(* IEC 61131-3 sources: STAR-PLC-Agent/results/raw/codex_matrix_resume_20261114/codex_deepseek/PUB012/functional/attempt_0001, 1 file *)

(* ---- test_program.st ---- *)
PROGRAM PLC_PRG
VAR
 BenchStep : UDINT := 0;
 BenchCalls : UDINT := 0;
 BenchDone : BOOL := FALSE;
 BenchLastTime : TIME := T#0ms;
 BenchClockReady : BOOL := FALSE;
 BenchCurrentTime : TIME := T#0ms;
 TraceDt : ARRAY[0..69] OF UDINT;
 BenchUut0 : FB_Task;
 BenchUut1 : FB_Task;
 BenchUut2 : FB_Task;
 BenchUut3 : FB_Task;
 BenchUut4 : FB_Task;
 BenchUut5 : FB_Task;
 BenchUut6 : FB_Task;
 BenchUut7 : FB_Task;
 TraceIn_THICKNESS_FAULT : ARRAY[0..69] OF BOOL;
 TraceIn_THICKNESS_SIGNAL_VALID : ARRAY[0..69] OF BOOL;
 TraceIn_CUTTING_RUN : ARRAY[0..69] OF BOOL;
 TraceIn_FaultTimestamp : ARRAY[0..69] OF DINT;
 TraceIn_CycleTime : ARRAY[0..69] OF TIME;
 TraceOut_THICKNESS_ALARM : ARRAY[0..69] OF BOOL;
 TraceOut_Slab_Fault_Counter : ARRAY[0..69] OF UINT;
 TraceOut_Slab_Runtime_Accumulator : ARRAY[0..69] OF LTIME;
 TraceOut_Slab_Fault_History_0 : ARRAY[0..69] OF DINT;
 TraceOut_Slab_Fault_History_1 : ARRAY[0..69] OF DINT;
 TraceOut_Slab_Fault_History_2 : ARRAY[0..69] OF DINT;
 TraceOut_Slab_Fault_History_3 : ARRAY[0..69] OF DINT;
 TraceOut_Slab_Fault_History_4 : ARRAY[0..69] OF DINT;
END_VAR

IF NOT BenchDone THEN
 BenchCurrentTime := TIME();
 IF NOT BenchClockReady THEN
  BenchLastTime := BenchCurrentTime;
  BenchClockReady := TRUE;
 ELSE
 CASE BenchStep OF
 0:
  IF BenchCurrentTime - BenchLastTime >= UDINT_TO_TIME(0) THEN
   TraceDt[0] := TIME_TO_UDINT(BenchCurrentTime - BenchLastTime);
   BenchLastTime := BenchCurrentTime;
   BenchUut0.THICKNESS_FAULT := FALSE;
   BenchUut0.THICKNESS_SIGNAL_VALID := TRUE;
   BenchUut0.CUTTING_RUN := FALSE;
   BenchUut0.FaultTimestamp := DINT#0;
   BenchUut0.CycleTime := T#100ms;
   TraceIn_THICKNESS_FAULT[0] := BenchUut0.THICKNESS_FAULT;
   TraceIn_THICKNESS_SIGNAL_VALID[0] := BenchUut0.THICKNESS_SIGNAL_VALID;
   TraceIn_CUTTING_RUN[0] := BenchUut0.CUTTING_RUN;
   TraceIn_FaultTimestamp[0] := BenchUut0.FaultTimestamp;
   TraceIn_CycleTime[0] := BenchUut0.CycleTime;
   BenchUut0();
   TraceOut_THICKNESS_ALARM[0] := BenchUut0.THICKNESS_ALARM;
   TraceOut_Slab_Fault_Counter[0] := BenchUut0.Slab_Fault_Counter;
   TraceOut_Slab_Runtime_Accumulator[0] := BenchUut0.Slab_Runtime_Accumulator;
   TraceOut_Slab_Fault_History_0[0] := BenchUut0.Slab_Fault_History[0];
   TraceOut_Slab_Fault_History_1[0] := BenchUut0.Slab_Fault_History[1];
   TraceOut_Slab_Fault_History_2[0] := BenchUut0.Slab_Fault_History[2];
   TraceOut_Slab_Fault_History_3[0] := BenchUut0.Slab_Fault_History[3];
   TraceOut_Slab_Fault_History_4[0] := BenchUut0.Slab_Fault_History[4];
   BenchCalls := BenchCalls + 1;
   BenchStep := BenchStep + 1;
  END_IF;
 1:
  IF BenchCurrentTime - BenchLastTime >= UDINT_TO_TIME(100) THEN
   TraceDt[1] := TIME_TO_UDINT(BenchCurrentTime - BenchLastTime);
   BenchLastTime := BenchCurrentTime;
   BenchUut0.THICKNESS_FAULT := TRUE;
   BenchUut0.THICKNESS_SIGNAL_VALID := TRUE;
   BenchUut0.CUTTING_RUN := FALSE;
   BenchUut0.FaultTimestamp := DINT#101;
   BenchUut0.CycleTime := T#100ms;
   TraceIn_THICKNESS_FAULT[1] := BenchUut0.THICKNESS_FAULT;
   TraceIn_THICKNESS_SIGNAL_VALID[1] := BenchUut0.THICKNESS_SIGNAL_VALID;
   TraceIn_CUTTING_RUN[1] := BenchUut0.CUTTING_RUN;
   TraceIn_FaultTimestamp[1] := BenchUut0.FaultTimestamp;
   TraceIn_CycleTime[1] := BenchUut0.CycleTime;
   BenchUut0();
   TraceOut_THICKNESS_ALARM[1] := BenchUut0.THICKNESS_ALARM;
   TraceOut_Slab_Fault_Counter[1] := BenchUut0.Slab_Fault_Counter;
   TraceOut_Slab_Runtime_Accumulator[1] := BenchUut0.Slab_Runtime_Accumulator;
   TraceOut_Slab_Fault_History_0[1] := BenchUut0.Slab_Fault_History[0];
   TraceOut_Slab_Fault_History_1[1] := BenchUut0.Slab_Fault_History[1];
   TraceOut_Slab_Fault_History_2[1] := BenchUut0.Slab_Fault_History[2];
   TraceOut_Slab_Fault_History_3[1] := BenchUut0.Slab_Fault_History[3];
   TraceOut_Slab_Fault_History_4[1] := BenchUut0.Slab_Fault_History[4];
   BenchCalls := BenchCalls + 1;
   BenchStep := BenchStep + 1;
  END_IF;
 2:
  IF BenchCurrentTime - BenchLastTime >= UDINT_TO_TIME(100) THEN
   TraceDt[2] := TIME_TO_UDINT(BenchCurrentTime - BenchLastTime);
   BenchLastTime := BenchCurrentTime;
   BenchUut0.THICKNESS_FAULT := FALSE;
   BenchUut0.THICKNESS_SIGNAL_VALID := TRUE;
   BenchUut0.CUTTING_RUN := FALSE;
   BenchUut0.FaultTimestamp := DINT#0;
   BenchUut0.CycleTime := T#100ms;
   TraceIn_THICKNESS_FAULT[2] := BenchUut0.THICKNESS_FAULT;
   TraceIn_THICKNESS_SIGNAL_VALID[2] := BenchUut0.THICKNESS_SIGNAL_VALID;
   TraceIn_CUTTING_RUN[2] := BenchUut0.CUTTING_RUN;
   TraceIn_FaultTimestamp[2] := BenchUut0.FaultTimestamp;
   TraceIn_CycleTime[2] := BenchUut0.CycleTime;
   BenchUut0();
   TraceOut_THICKNESS_ALARM[2] := BenchUut0.THICKNESS_ALARM;
   TraceOut_Slab_Fault_Counter[2] := BenchUut0.Slab_Fault_Counter;
   TraceOut_Slab_Runtime_Accumulator[2] := BenchUut0.Slab_Runtime_Accumulator;
   TraceOut_Slab_Fault_History_0[2] := BenchUut0.Slab_Fault_History[0];
   TraceOut_Slab_Fault_History_1[2] := BenchUut0.Slab_Fault_History[1];
   TraceOut_Slab_Fault_History_2[2] := BenchUut0.Slab_Fault_History[2];
   TraceOut_Slab_Fault_History_3[2] := BenchUut0.Slab_Fault_History[3];
   TraceOut_Slab_Fault_History_4[2] := BenchUut0.Slab_Fault_History[4];
   BenchCalls := BenchCalls + 1;
   BenchStep := BenchStep + 1;
  END_IF;
 3:
  IF BenchCurrentTime - BenchLastTime >= UDINT_TO_TIME(300) THEN
   TraceDt[3] := TIME_TO_UDINT(BenchCurrentTime - BenchLastTime);
   BenchLastTime := BenchCurrentTime;
   BenchUut0.THICKNESS_FAULT := FALSE;
   BenchUut0.THICKNESS_SIGNAL_VALID := TRUE;
   BenchUut0.CUTTING_RUN := FALSE;
   BenchUut0.FaultTimestamp := DINT#0;
   BenchUut0.CycleTime := T#100ms;
   TraceIn_THICKNESS_FAULT[3] := BenchUut0.THICKNESS_FAULT;
   TraceIn_THICKNESS_SIGNAL_VALID[3] := BenchUut0.THICKNESS_SIGNAL_VALID;
   TraceIn_CUTTING_RUN[3] := BenchUut0.CUTTING_RUN;
   TraceIn_FaultTimestamp[3] := BenchUut0.FaultTimestamp;
   TraceIn_CycleTime[3] := BenchUut0.CycleTime;
   BenchUut0();
   TraceOut_THICKNESS_ALARM[3] := BenchUut0.THICKNESS_ALARM;
   TraceOut_Slab_Fault_Counter[3] := BenchUut0.Slab_Fault_Counter;
   TraceOut_Slab_Runtime_Accumulator[3] := BenchUut0.Slab_Runtime_Accumulator;
   TraceOut_Slab_Fault_History_0[3] := BenchUut0.Slab_Fault_History[0];
   TraceOut_Slab_Fault_History_1[3] := BenchUut0.Slab_Fault_History[1];
   TraceOut_Slab_Fault_History_2[3] := BenchUut0.Slab_Fault_History[2];
   TraceOut_Slab_Fault_History_3[3] := BenchUut0.Slab_Fault_History[3];
   TraceOut_Slab_Fault_History_4[3] := BenchUut0.Slab_Fault_History[4];
   BenchCalls := BenchCalls + 1;
   BenchStep := BenchStep + 1;
  END_IF;
 4:
  IF BenchCurrentTime - BenchLastTime >= UDINT_TO_TIME(100) THEN
   TraceDt[4] := TIME_TO_UDINT(BenchCurrentTime - BenchLastTime);
   BenchLastTime := BenchCurrentTime;
   BenchUut0.THICKNESS_FAULT := FALSE;
   BenchUut0.THICKNESS_SIGNAL_VALID := TRUE;
   BenchUut0.CUTTING_RUN := FALSE;
   BenchUut0.FaultTimestamp := DINT#0;
   BenchUut0.CycleTime := T#100ms;
   TraceIn_THICKNESS_FAULT[4] := BenchUut0.THICKNESS_FAULT;
   TraceIn_THICKNESS_SIGNAL_VALID[4] := BenchUut0.THICKNESS_SIGNAL_VALID;
   TraceIn_CUTTING_RUN[4] := BenchUut0.CUTTING_RUN;
   TraceIn_FaultTimestamp[4] := BenchUut0.FaultTimestamp;
   TraceIn_CycleTime[4] := BenchUut0.CycleTime;
   BenchUut0();
   TraceOut_THICKNESS_ALARM[4] := BenchUut0.THICKNESS_ALARM;
   TraceOut_Slab_Fault_Counter[4] := BenchUut0.Slab_Fault_Counter;
   TraceOut_Slab_Runtime_Accumulator[4] := BenchUut0.Slab_Runtime_Accumulator;
   TraceOut_Slab_Fault_History_0[4] := BenchUut0.Slab_Fault_History[0];
   TraceOut_Slab_Fault_History_1[4] := BenchUut0.Slab_Fault_History[1];
   TraceOut_Slab_Fault_History_2[4] := BenchUut0.Slab_Fault_History[2];
   TraceOut_Slab_Fault_History_3[4] := BenchUut0.Slab_Fault_History[3];
   TraceOut_Slab_Fault_History_4[4] := BenchUut0.Slab_Fault_History[4];
   BenchCalls := BenchCalls + 1;
   BenchStep := BenchStep + 1;
  END_IF;
 5:
  IF BenchCurrentTime - BenchLastTime >= UDINT_TO_TIME(100) THEN
   TraceDt[5] := TIME_TO_UDINT(BenchCurrentTime - BenchLastTime);
   BenchLastTime := BenchCurrentTime;
   BenchUut0.THICKNESS_FAULT := TRUE;
   BenchUut0.THICKNESS_SIGNAL_VALID := TRUE;
   BenchUut0.CUTTING_RUN := FALSE;
   BenchUut0.FaultTimestamp := DINT#102;
   BenchUut0.CycleTime := T#100ms;
   TraceIn_THICKNESS_FAULT[5] := BenchUut0.THICKNESS_FAULT;
   TraceIn_THICKNESS_SIGNAL_VALID[5] := BenchUut0.THICKNESS_SIGNAL_VALID;
   TraceIn_CUTTING_RUN[5] := BenchUut0.CUTTING_RUN;
   TraceIn_FaultTimestamp[5] := BenchUut0.FaultTimestamp;
   TraceIn_CycleTime[5] := BenchUut0.CycleTime;
   BenchUut0();
   TraceOut_THICKNESS_ALARM[5] := BenchUut0.THICKNESS_ALARM;
   TraceOut_Slab_Fault_Counter[5] := BenchUut0.Slab_Fault_Counter;
   TraceOut_Slab_Runtime_Accumulator[5] := BenchUut0.Slab_Runtime_Accumulator;
   TraceOut_Slab_Fault_History_0[5] := BenchUut0.Slab_Fault_History[0];
   TraceOut_Slab_Fault_History_1[5] := BenchUut0.Slab_Fault_History[1];
   TraceOut_Slab_Fault_History_2[5] := BenchUut0.Slab_Fault_History[2];
   TraceOut_Slab_Fault_History_3[5] := BenchUut0.Slab_Fault_History[3];
   TraceOut_Slab_Fault_History_4[5] := BenchUut0.Slab_Fault_History[4];
   BenchCalls := BenchCalls + 1;
   BenchStep := BenchStep + 1;
  END_IF;
 6:
  IF BenchCurrentTime - BenchLastTime >= UDINT_TO_TIME(10) THEN
   TraceDt[6] := TIME_TO_UDINT(BenchCurrentTime - BenchLastTime);
   BenchLastTime := BenchCurrentTime;
   BenchUut0.THICKNESS_FAULT := TRUE;
   BenchUut0.THICKNESS_SIGNAL_VALID := FALSE;
   BenchUut0.CUTTING_RUN := FALSE;
   BenchUut0.FaultTimestamp := DINT#0;
   BenchUut0.CycleTime := T#100ms;
   TraceIn_THICKNESS_FAULT[6] := BenchUut0.THICKNESS_FAULT;
   TraceIn_THICKNESS_SIGNAL_VALID[6] := BenchUut0.THICKNESS_SIGNAL_VALID;
   TraceIn_CUTTING_RUN[6] := BenchUut0.CUTTING_RUN;
   TraceIn_FaultTimestamp[6] := BenchUut0.FaultTimestamp;
   TraceIn_CycleTime[6] := BenchUut0.CycleTime;
   BenchUut0();
   TraceOut_THICKNESS_ALARM[6] := BenchUut0.THICKNESS_ALARM;
   TraceOut_Slab_Fault_Counter[6] := BenchUut0.Slab_Fault_Counter;
   TraceOut_Slab_Runtime_Accumulator[6] := BenchUut0.Slab_Runtime_Accumulator;
   TraceOut_Slab_Fault_History_0[6] := BenchUut0.Slab_Fault_History[0];
   TraceOut_Slab_Fault_History_1[6] := BenchUut0.Slab_Fault_History[1];
   TraceOut_Slab_Fault_History_2[6] := BenchUut0.Slab_Fault_History[2];
   TraceOut_Slab_Fault_History_3[6] := BenchUut0.Slab_Fault_History[3];
   TraceOut_Slab_Fault_History_4[6] := BenchUut0.Slab_Fault_History[4];
   BenchCalls := BenchCalls + 1;
   BenchStep := BenchStep + 1;
  END_IF;
 7:
  IF BenchCurrentTime - BenchLastTime >= UDINT_TO_TIME(0) THEN
   TraceDt[7] := TIME_TO_UDINT(BenchCurrentTime - BenchLastTime);
   BenchLastTime := BenchCurrentTime;
   BenchUut1.THICKNESS_FAULT := FALSE;
   BenchUut1.THICKNESS_SIGNAL_VALID := TRUE;
   BenchUut1.CUTTING_RUN := FALSE;
   BenchUut1.FaultTimestamp := DINT#0;
   BenchUut1.CycleTime := T#100ms;
   TraceIn_THICKNESS_FAULT[7] := BenchUut1.THICKNESS_FAULT;
   TraceIn_THICKNESS_SIGNAL_VALID[7] := BenchUut1.THICKNESS_SIGNAL_VALID;
   TraceIn_CUTTING_RUN[7] := BenchUut1.CUTTING_RUN;
   TraceIn_FaultTimestamp[7] := BenchUut1.FaultTimestamp;
   TraceIn_CycleTime[7] := BenchUut1.CycleTime;
   BenchUut1();
   TraceOut_THICKNESS_ALARM[7] := BenchUut1.THICKNESS_ALARM;
   TraceOut_Slab_Fault_Counter[7] := BenchUut1.Slab_Fault_Counter;
   TraceOut_Slab_Runtime_Accumulator[7] := BenchUut1.Slab_Runtime_Accumulator;
   TraceOut_Slab_Fault_History_0[7] := BenchUut1.Slab_Fault_History[0];
   TraceOut_Slab_Fault_History_1[7] := BenchUut1.Slab_Fault_History[1];
   TraceOut_Slab_Fault_History_2[7] := BenchUut1.Slab_Fault_History[2];
   TraceOut_Slab_Fault_History_3[7] := BenchUut1.Slab_Fault_History[3];
   TraceOut_Slab_Fault_History_4[7] := BenchUut1.Slab_Fault_History[4];
   BenchCalls := BenchCalls + 1;
   BenchStep := BenchStep + 1;
  END_IF;
 8:
  IF BenchCurrentTime - BenchLastTime >= UDINT_TO_TIME(100) THEN
   TraceDt[8] := TIME_TO_UDINT(BenchCurrentTime - BenchLastTime);
   BenchLastTime := BenchCurrentTime;
   BenchUut1.THICKNESS_FAULT := TRUE;
   BenchUut1.THICKNESS_SIGNAL_VALID := TRUE;
   BenchUut1.CUTTING_RUN := FALSE;
   BenchUut1.FaultTimestamp := DINT#1;
   BenchUut1.CycleTime := T#100ms;
   TraceIn_THICKNESS_FAULT[8] := BenchUut1.THICKNESS_FAULT;
   TraceIn_THICKNESS_SIGNAL_VALID[8] := BenchUut1.THICKNESS_SIGNAL_VALID;
   TraceIn_CUTTING_RUN[8] := BenchUut1.CUTTING_RUN;
   TraceIn_FaultTimestamp[8] := BenchUut1.FaultTimestamp;
   TraceIn_CycleTime[8] := BenchUut1.CycleTime;
   BenchUut1();
   TraceOut_THICKNESS_ALARM[8] := BenchUut1.THICKNESS_ALARM;
   TraceOut_Slab_Fault_Counter[8] := BenchUut1.Slab_Fault_Counter;
   TraceOut_Slab_Runtime_Accumulator[8] := BenchUut1.Slab_Runtime_Accumulator;
   TraceOut_Slab_Fault_History_0[8] := BenchUut1.Slab_Fault_History[0];
   TraceOut_Slab_Fault_History_1[8] := BenchUut1.Slab_Fault_History[1];
   TraceOut_Slab_Fault_History_2[8] := BenchUut1.Slab_Fault_History[2];
   TraceOut_Slab_Fault_History_3[8] := BenchUut1.Slab_Fault_History[3];
   TraceOut_Slab_Fault_History_4[8] := BenchUut1.Slab_Fault_History[4];
   BenchCalls := BenchCalls + 1;
   BenchStep := BenchStep + 1;
  END_IF;
 9:
  IF BenchCurrentTime - BenchLastTime >= UDINT_TO_TIME(100) THEN
   TraceDt[9] := TIME_TO_UDINT(BenchCurrentTime - BenchLastTime);
   BenchLastTime := BenchCurrentTime;
   BenchUut1.THICKNESS_FAULT := FALSE;
   BenchUut1.THICKNESS_SIGNAL_VALID := TRUE;
   BenchUut1.CUTTING_RUN := FALSE;
   BenchUut1.FaultTimestamp := DINT#0;
   BenchUut1.CycleTime := T#100ms;
   TraceIn_THICKNESS_FAULT[9] := BenchUut1.THICKNESS_FAULT;
   TraceIn_THICKNESS_SIGNAL_VALID[9] := BenchUut1.THICKNESS_SIGNAL_VALID;
   TraceIn_CUTTING_RUN[9] := BenchUut1.CUTTING_RUN;
   TraceIn_FaultTimestamp[9] := BenchUut1.FaultTimestamp;
   TraceIn_CycleTime[9] := BenchUut1.CycleTime;
   BenchUut1();
   TraceOut_THICKNESS_ALARM[9] := BenchUut1.THICKNESS_ALARM;
   TraceOut_Slab_Fault_Counter[9] := BenchUut1.Slab_Fault_Counter;
   TraceOut_Slab_Runtime_Accumulator[9] := BenchUut1.Slab_Runtime_Accumulator;
   TraceOut_Slab_Fault_History_0[9] := BenchUut1.Slab_Fault_History[0];
   TraceOut_Slab_Fault_History_1[9] := BenchUut1.Slab_Fault_History[1];
   TraceOut_Slab_Fault_History_2[9] := BenchUut1.Slab_Fault_History[2];
   TraceOut_Slab_Fault_History_3[9] := BenchUut1.Slab_Fault_History[3];
   TraceOut_Slab_Fault_History_4[9] := BenchUut1.Slab_Fault_History[4];
   BenchCalls := BenchCalls + 1;
   BenchStep := BenchStep + 1;
  END_IF;
 10:
  IF BenchCurrentTime - BenchLastTime >= UDINT_TO_TIME(100) THEN
   TraceDt[10] := TIME_TO_UDINT(BenchCurrentTime - BenchLastTime);
   BenchLastTime := BenchCurrentTime;
   BenchUut1.THICKNESS_FAULT := TRUE;
   BenchUut1.THICKNESS_SIGNAL_VALID := TRUE;
   BenchUut1.CUTTING_RUN := FALSE;
   BenchUut1.FaultTimestamp := DINT#2;
   BenchUut1.CycleTime := T#100ms;
   TraceIn_THICKNESS_FAULT[10] := BenchUut1.THICKNESS_FAULT;
   TraceIn_THICKNESS_SIGNAL_VALID[10] := BenchUut1.THICKNESS_SIGNAL_VALID;
   TraceIn_CUTTING_RUN[10] := BenchUut1.CUTTING_RUN;
   TraceIn_FaultTimestamp[10] := BenchUut1.FaultTimestamp;
   TraceIn_CycleTime[10] := BenchUut1.CycleTime;
   BenchUut1();
   TraceOut_THICKNESS_ALARM[10] := BenchUut1.THICKNESS_ALARM;
   TraceOut_Slab_Fault_Counter[10] := BenchUut1.Slab_Fault_Counter;
   TraceOut_Slab_Runtime_Accumulator[10] := BenchUut1.Slab_Runtime_Accumulator;
   TraceOut_Slab_Fault_History_0[10] := BenchUut1.Slab_Fault_History[0];
   TraceOut_Slab_Fault_History_1[10] := BenchUut1.Slab_Fault_History[1];
   TraceOut_Slab_Fault_History_2[10] := BenchUut1.Slab_Fault_History[2];
   TraceOut_Slab_Fault_History_3[10] := BenchUut1.Slab_Fault_History[3];
   TraceOut_Slab_Fault_History_4[10] := BenchUut1.Slab_Fault_History[4];
   BenchCalls := BenchCalls + 1;
   BenchStep := BenchStep + 1;
  END_IF;
 11:
  IF BenchCurrentTime - BenchLastTime >= UDINT_TO_TIME(100) THEN
   TraceDt[11] := TIME_TO_UDINT(BenchCurrentTime - BenchLastTime);
   BenchLastTime := BenchCurrentTime;
   BenchUut1.THICKNESS_FAULT := FALSE;
   BenchUut1.THICKNESS_SIGNAL_VALID := TRUE;
   BenchUut1.CUTTING_RUN := FALSE;
   BenchUut1.FaultTimestamp := DINT#0;
   BenchUut1.CycleTime := T#100ms;
   TraceIn_THICKNESS_FAULT[11] := BenchUut1.THICKNESS_FAULT;
   TraceIn_THICKNESS_SIGNAL_VALID[11] := BenchUut1.THICKNESS_SIGNAL_VALID;
   TraceIn_CUTTING_RUN[11] := BenchUut1.CUTTING_RUN;
   TraceIn_FaultTimestamp[11] := BenchUut1.FaultTimestamp;
   TraceIn_CycleTime[11] := BenchUut1.CycleTime;
   BenchUut1();
   TraceOut_THICKNESS_ALARM[11] := BenchUut1.THICKNESS_ALARM;
   TraceOut_Slab_Fault_Counter[11] := BenchUut1.Slab_Fault_Counter;
   TraceOut_Slab_Runtime_Accumulator[11] := BenchUut1.Slab_Runtime_Accumulator;
   TraceOut_Slab_Fault_History_0[11] := BenchUut1.Slab_Fault_History[0];
   TraceOut_Slab_Fault_History_1[11] := BenchUut1.Slab_Fault_History[1];
   TraceOut_Slab_Fault_History_2[11] := BenchUut1.Slab_Fault_History[2];
   TraceOut_Slab_Fault_History_3[11] := BenchUut1.Slab_Fault_History[3];
   TraceOut_Slab_Fault_History_4[11] := BenchUut1.Slab_Fault_History[4];
   BenchCalls := BenchCalls + 1;
   BenchStep := BenchStep + 1;
  END_IF;
 12:
  IF BenchCurrentTime - BenchLastTime >= UDINT_TO_TIME(100) THEN
   TraceDt[12] := TIME_TO_UDINT(BenchCurrentTime - BenchLastTime);
   BenchLastTime := BenchCurrentTime;
   BenchUut1.THICKNESS_FAULT := TRUE;
   BenchUut1.THICKNESS_SIGNAL_VALID := TRUE;
   BenchUut1.CUTTING_RUN := FALSE;
   BenchUut1.FaultTimestamp := DINT#3;
   BenchUut1.CycleTime := T#100ms;
   TraceIn_THICKNESS_FAULT[12] := BenchUut1.THICKNESS_FAULT;
   TraceIn_THICKNESS_SIGNAL_VALID[12] := BenchUut1.THICKNESS_SIGNAL_VALID;
   TraceIn_CUTTING_RUN[12] := BenchUut1.CUTTING_RUN;
   TraceIn_FaultTimestamp[12] := BenchUut1.FaultTimestamp;
   TraceIn_CycleTime[12] := BenchUut1.CycleTime;
   BenchUut1();
   TraceOut_THICKNESS_ALARM[12] := BenchUut1.THICKNESS_ALARM;
   TraceOut_Slab_Fault_Counter[12] := BenchUut1.Slab_Fault_Counter;
   TraceOut_Slab_Runtime_Accumulator[12] := BenchUut1.Slab_Runtime_Accumulator;
   TraceOut_Slab_Fault_History_0[12] := BenchUut1.Slab_Fault_History[0];
   TraceOut_Slab_Fault_History_1[12] := BenchUut1.Slab_Fault_History[1];
   TraceOut_Slab_Fault_History_2[12] := BenchUut1.Slab_Fault_History[2];
   TraceOut_Slab_Fault_History_3[12] := BenchUut1.Slab_Fault_History[3];
   TraceOut_Slab_Fault_History_4[12] := BenchUut1.Slab_Fault_History[4];
   BenchCalls := BenchCalls + 1;
   BenchStep := BenchStep + 1;
  END_IF;
 13:
  IF BenchCurrentTime - BenchLastTime >= UDINT_TO_TIME(100) THEN
   TraceDt[13] := TIME_TO_UDINT(BenchCurrentTime - BenchLastTime);
   BenchLastTime := BenchCurrentTime;
   BenchUut1.THICKNESS_FAULT := FALSE;
   BenchUut1.THICKNESS_SIGNAL_VALID := TRUE;
   BenchUut1.CUTTING_RUN := FALSE;
   BenchUut1.FaultTimestamp := DINT#0;
   BenchUut1.CycleTime := T#100ms;
   TraceIn_THICKNESS_FAULT[13] := BenchUut1.THICKNESS_FAULT;
   TraceIn_THICKNESS_SIGNAL_VALID[13] := BenchUut1.THICKNESS_SIGNAL_VALID;
   TraceIn_CUTTING_RUN[13] := BenchUut1.CUTTING_RUN;
   TraceIn_FaultTimestamp[13] := BenchUut1.FaultTimestamp;
   TraceIn_CycleTime[13] := BenchUut1.CycleTime;
   BenchUut1();
   TraceOut_THICKNESS_ALARM[13] := BenchUut1.THICKNESS_ALARM;
   TraceOut_Slab_Fault_Counter[13] := BenchUut1.Slab_Fault_Counter;
   TraceOut_Slab_Runtime_Accumulator[13] := BenchUut1.Slab_Runtime_Accumulator;
   TraceOut_Slab_Fault_History_0[13] := BenchUut1.Slab_Fault_History[0];
   TraceOut_Slab_Fault_History_1[13] := BenchUut1.Slab_Fault_History[1];
   TraceOut_Slab_Fault_History_2[13] := BenchUut1.Slab_Fault_History[2];
   TraceOut_Slab_Fault_History_3[13] := BenchUut1.Slab_Fault_History[3];
   TraceOut_Slab_Fault_History_4[13] := BenchUut1.Slab_Fault_History[4];
   BenchCalls := BenchCalls + 1;
   BenchStep := BenchStep + 1;
  END_IF;
 14:
  IF BenchCurrentTime - BenchLastTime >= UDINT_TO_TIME(100) THEN
   TraceDt[14] := TIME_TO_UDINT(BenchCurrentTime - BenchLastTime);
   BenchLastTime := BenchCurrentTime;
   BenchUut1.THICKNESS_FAULT := TRUE;
   BenchUut1.THICKNESS_SIGNAL_VALID := TRUE;
   BenchUut1.CUTTING_RUN := FALSE;
   BenchUut1.FaultTimestamp := DINT#4;
   BenchUut1.CycleTime := T#100ms;
   TraceIn_THICKNESS_FAULT[14] := BenchUut1.THICKNESS_FAULT;
   TraceIn_THICKNESS_SIGNAL_VALID[14] := BenchUut1.THICKNESS_SIGNAL_VALID;
   TraceIn_CUTTING_RUN[14] := BenchUut1.CUTTING_RUN;
   TraceIn_FaultTimestamp[14] := BenchUut1.FaultTimestamp;
   TraceIn_CycleTime[14] := BenchUut1.CycleTime;
   BenchUut1();
   TraceOut_THICKNESS_ALARM[14] := BenchUut1.THICKNESS_ALARM;
   TraceOut_Slab_Fault_Counter[14] := BenchUut1.Slab_Fault_Counter;
   TraceOut_Slab_Runtime_Accumulator[14] := BenchUut1.Slab_Runtime_Accumulator;
   TraceOut_Slab_Fault_History_0[14] := BenchUut1.Slab_Fault_History[0];
   TraceOut_Slab_Fault_History_1[14] := BenchUut1.Slab_Fault_History[1];
   TraceOut_Slab_Fault_History_2[14] := BenchUut1.Slab_Fault_History[2];
   TraceOut_Slab_Fault_History_3[14] := BenchUut1.Slab_Fault_History[3];
   TraceOut_Slab_Fault_History_4[14] := BenchUut1.Slab_Fault_History[4];
   BenchCalls := BenchCalls + 1;
   BenchStep := BenchStep + 1;
  END_IF;
 15:
  IF BenchCurrentTime - BenchLastTime >= UDINT_TO_TIME(100) THEN
   TraceDt[15] := TIME_TO_UDINT(BenchCurrentTime - BenchLastTime);
   BenchLastTime := BenchCurrentTime;
   BenchUut1.THICKNESS_FAULT := FALSE;
   BenchUut1.THICKNESS_SIGNAL_VALID := TRUE;
   BenchUut1.CUTTING_RUN := FALSE;
   BenchUut1.FaultTimestamp := DINT#0;
   BenchUut1.CycleTime := T#100ms;
   TraceIn_THICKNESS_FAULT[15] := BenchUut1.THICKNESS_FAULT;
   TraceIn_THICKNESS_SIGNAL_VALID[15] := BenchUut1.THICKNESS_SIGNAL_VALID;
   TraceIn_CUTTING_RUN[15] := BenchUut1.CUTTING_RUN;
   TraceIn_FaultTimestamp[15] := BenchUut1.FaultTimestamp;
   TraceIn_CycleTime[15] := BenchUut1.CycleTime;
   BenchUut1();
   TraceOut_THICKNESS_ALARM[15] := BenchUut1.THICKNESS_ALARM;
   TraceOut_Slab_Fault_Counter[15] := BenchUut1.Slab_Fault_Counter;
   TraceOut_Slab_Runtime_Accumulator[15] := BenchUut1.Slab_Runtime_Accumulator;
   TraceOut_Slab_Fault_History_0[15] := BenchUut1.Slab_Fault_History[0];
   TraceOut_Slab_Fault_History_1[15] := BenchUut1.Slab_Fault_History[1];
   TraceOut_Slab_Fault_History_2[15] := BenchUut1.Slab_Fault_History[2];
   TraceOut_Slab_Fault_History_3[15] := BenchUut1.Slab_Fault_History[3];
   TraceOut_Slab_Fault_History_4[15] := BenchUut1.Slab_Fault_History[4];
   BenchCalls := BenchCalls + 1;
   BenchStep := BenchStep + 1;
  END_IF;
 16:
  IF BenchCurrentTime - BenchLastTime >= UDINT_TO_TIME(100) THEN
   TraceDt[16] := TIME_TO_UDINT(BenchCurrentTime - BenchLastTime);
   BenchLastTime := BenchCurrentTime;
   BenchUut1.THICKNESS_FAULT := TRUE;
   BenchUut1.THICKNESS_SIGNAL_VALID := TRUE;
   BenchUut1.CUTTING_RUN := FALSE;
   BenchUut1.FaultTimestamp := DINT#5;
   BenchUut1.CycleTime := T#100ms;
   TraceIn_THICKNESS_FAULT[16] := BenchUut1.THICKNESS_FAULT;
   TraceIn_THICKNESS_SIGNAL_VALID[16] := BenchUut1.THICKNESS_SIGNAL_VALID;
   TraceIn_CUTTING_RUN[16] := BenchUut1.CUTTING_RUN;
   TraceIn_FaultTimestamp[16] := BenchUut1.FaultTimestamp;
   TraceIn_CycleTime[16] := BenchUut1.CycleTime;
   BenchUut1();
   TraceOut_THICKNESS_ALARM[16] := BenchUut1.THICKNESS_ALARM;
   TraceOut_Slab_Fault_Counter[16] := BenchUut1.Slab_Fault_Counter;
   TraceOut_Slab_Runtime_Accumulator[16] := BenchUut1.Slab_Runtime_Accumulator;
   TraceOut_Slab_Fault_History_0[16] := BenchUut1.Slab_Fault_History[0];
   TraceOut_Slab_Fault_History_1[16] := BenchUut1.Slab_Fault_History[1];
   TraceOut_Slab_Fault_History_2[16] := BenchUut1.Slab_Fault_History[2];
   TraceOut_Slab_Fault_History_3[16] := BenchUut1.Slab_Fault_History[3];
   TraceOut_Slab_Fault_History_4[16] := BenchUut1.Slab_Fault_History[4];
   BenchCalls := BenchCalls + 1;
   BenchStep := BenchStep + 1;
  END_IF;
 17:
  IF BenchCurrentTime - BenchLastTime >= UDINT_TO_TIME(100) THEN
   TraceDt[17] := TIME_TO_UDINT(BenchCurrentTime - BenchLastTime);
   BenchLastTime := BenchCurrentTime;
   BenchUut1.THICKNESS_FAULT := FALSE;
   BenchUut1.THICKNESS_SIGNAL_VALID := TRUE;
   BenchUut1.CUTTING_RUN := FALSE;
   BenchUut1.FaultTimestamp := DINT#0;
   BenchUut1.CycleTime := T#100ms;
   TraceIn_THICKNESS_FAULT[17] := BenchUut1.THICKNESS_FAULT;
   TraceIn_THICKNESS_SIGNAL_VALID[17] := BenchUut1.THICKNESS_SIGNAL_VALID;
   TraceIn_CUTTING_RUN[17] := BenchUut1.CUTTING_RUN;
   TraceIn_FaultTimestamp[17] := BenchUut1.FaultTimestamp;
   TraceIn_CycleTime[17] := BenchUut1.CycleTime;
   BenchUut1();
   TraceOut_THICKNESS_ALARM[17] := BenchUut1.THICKNESS_ALARM;
   TraceOut_Slab_Fault_Counter[17] := BenchUut1.Slab_Fault_Counter;
   TraceOut_Slab_Runtime_Accumulator[17] := BenchUut1.Slab_Runtime_Accumulator;
   TraceOut_Slab_Fault_History_0[17] := BenchUut1.Slab_Fault_History[0];
   TraceOut_Slab_Fault_History_1[17] := BenchUut1.Slab_Fault_History[1];
   TraceOut_Slab_Fault_History_2[17] := BenchUut1.Slab_Fault_History[2];
   TraceOut_Slab_Fault_History_3[17] := BenchUut1.Slab_Fault_History[3];
   TraceOut_Slab_Fault_History_4[17] := BenchUut1.Slab_Fault_History[4];
   BenchCalls := BenchCalls + 1;
   BenchStep := BenchStep + 1;
  END_IF;
 18:
  IF BenchCurrentTime - BenchLastTime >= UDINT_TO_TIME(100) THEN
   TraceDt[18] := TIME_TO_UDINT(BenchCurrentTime - BenchLastTime);
   BenchLastTime := BenchCurrentTime;
   BenchUut1.THICKNESS_FAULT := TRUE;
   BenchUut1.THICKNESS_SIGNAL_VALID := TRUE;
   BenchUut1.CUTTING_RUN := FALSE;
   BenchUut1.FaultTimestamp := DINT#6;
   BenchUut1.CycleTime := T#100ms;
   TraceIn_THICKNESS_FAULT[18] := BenchUut1.THICKNESS_FAULT;
   TraceIn_THICKNESS_SIGNAL_VALID[18] := BenchUut1.THICKNESS_SIGNAL_VALID;
   TraceIn_CUTTING_RUN[18] := BenchUut1.CUTTING_RUN;
   TraceIn_FaultTimestamp[18] := BenchUut1.FaultTimestamp;
   TraceIn_CycleTime[18] := BenchUut1.CycleTime;
   BenchUut1();
   TraceOut_THICKNESS_ALARM[18] := BenchUut1.THICKNESS_ALARM;
   TraceOut_Slab_Fault_Counter[18] := BenchUut1.Slab_Fault_Counter;
   TraceOut_Slab_Runtime_Accumulator[18] := BenchUut1.Slab_Runtime_Accumulator;
   TraceOut_Slab_Fault_History_0[18] := BenchUut1.Slab_Fault_History[0];
   TraceOut_Slab_Fault_History_1[18] := BenchUut1.Slab_Fault_History[1];
   TraceOut_Slab_Fault_History_2[18] := BenchUut1.Slab_Fault_History[2];
   TraceOut_Slab_Fault_History_3[18] := BenchUut1.Slab_Fault_History[3];
   TraceOut_Slab_Fault_History_4[18] := BenchUut1.Slab_Fault_History[4];
   BenchCalls := BenchCalls + 1;
   BenchStep := BenchStep + 1;
  END_IF;
 19:
  IF BenchCurrentTime - BenchLastTime >= UDINT_TO_TIME(100) THEN
   TraceDt[19] := TIME_TO_UDINT(BenchCurrentTime - BenchLastTime);
   BenchLastTime := BenchCurrentTime;
   BenchUut1.THICKNESS_FAULT := FALSE;
   BenchUut1.THICKNESS_SIGNAL_VALID := TRUE;
   BenchUut1.CUTTING_RUN := FALSE;
   BenchUut1.FaultTimestamp := DINT#0;
   BenchUut1.CycleTime := T#100ms;
   TraceIn_THICKNESS_FAULT[19] := BenchUut1.THICKNESS_FAULT;
   TraceIn_THICKNESS_SIGNAL_VALID[19] := BenchUut1.THICKNESS_SIGNAL_VALID;
   TraceIn_CUTTING_RUN[19] := BenchUut1.CUTTING_RUN;
   TraceIn_FaultTimestamp[19] := BenchUut1.FaultTimestamp;
   TraceIn_CycleTime[19] := BenchUut1.CycleTime;
   BenchUut1();
   TraceOut_THICKNESS_ALARM[19] := BenchUut1.THICKNESS_ALARM;
   TraceOut_Slab_Fault_Counter[19] := BenchUut1.Slab_Fault_Counter;
   TraceOut_Slab_Runtime_Accumulator[19] := BenchUut1.Slab_Runtime_Accumulator;
   TraceOut_Slab_Fault_History_0[19] := BenchUut1.Slab_Fault_History[0];
   TraceOut_Slab_Fault_History_1[19] := BenchUut1.Slab_Fault_History[1];
   TraceOut_Slab_Fault_History_2[19] := BenchUut1.Slab_Fault_History[2];
   TraceOut_Slab_Fault_History_3[19] := BenchUut1.Slab_Fault_History[3];
   TraceOut_Slab_Fault_History_4[19] := BenchUut1.Slab_Fault_History[4];
   BenchCalls := BenchCalls + 1;
   BenchStep := BenchStep + 1;
  END_IF;
 20:
  IF BenchCurrentTime - BenchLastTime >= UDINT_TO_TIME(0) THEN
   TraceDt[20] := TIME_TO_UDINT(BenchCurrentTime - BenchLastTime);
   BenchLastTime := BenchCurrentTime;
   BenchUut2.THICKNESS_FAULT := FALSE;
   BenchUut2.THICKNESS_SIGNAL_VALID := TRUE;
   BenchUut2.CUTTING_RUN := TRUE;
   BenchUut2.FaultTimestamp := DINT#0;
   BenchUut2.CycleTime := T#100ms;
   TraceIn_THICKNESS_FAULT[20] := BenchUut2.THICKNESS_FAULT;
   TraceIn_THICKNESS_SIGNAL_VALID[20] := BenchUut2.THICKNESS_SIGNAL_VALID;
   TraceIn_CUTTING_RUN[20] := BenchUut2.CUTTING_RUN;
   TraceIn_FaultTimestamp[20] := BenchUut2.FaultTimestamp;
   TraceIn_CycleTime[20] := BenchUut2.CycleTime;
   BenchUut2();
   TraceOut_THICKNESS_ALARM[20] := BenchUut2.THICKNESS_ALARM;
   TraceOut_Slab_Fault_Counter[20] := BenchUut2.Slab_Fault_Counter;
   TraceOut_Slab_Runtime_Accumulator[20] := BenchUut2.Slab_Runtime_Accumulator;
   TraceOut_Slab_Fault_History_0[20] := BenchUut2.Slab_Fault_History[0];
   TraceOut_Slab_Fault_History_1[20] := BenchUut2.Slab_Fault_History[1];
   TraceOut_Slab_Fault_History_2[20] := BenchUut2.Slab_Fault_History[2];
   TraceOut_Slab_Fault_History_3[20] := BenchUut2.Slab_Fault_History[3];
   TraceOut_Slab_Fault_History_4[20] := BenchUut2.Slab_Fault_History[4];
   BenchCalls := BenchCalls + 1;
   BenchStep := BenchStep + 1;
  END_IF;
 21:
  IF BenchCurrentTime - BenchLastTime >= UDINT_TO_TIME(100) THEN
   TraceDt[21] := TIME_TO_UDINT(BenchCurrentTime - BenchLastTime);
   BenchLastTime := BenchCurrentTime;
   BenchUut2.THICKNESS_FAULT := FALSE;
   BenchUut2.THICKNESS_SIGNAL_VALID := TRUE;
   BenchUut2.CUTTING_RUN := TRUE;
   BenchUut2.FaultTimestamp := DINT#0;
   BenchUut2.CycleTime := T#100ms;
   TraceIn_THICKNESS_FAULT[21] := BenchUut2.THICKNESS_FAULT;
   TraceIn_THICKNESS_SIGNAL_VALID[21] := BenchUut2.THICKNESS_SIGNAL_VALID;
   TraceIn_CUTTING_RUN[21] := BenchUut2.CUTTING_RUN;
   TraceIn_FaultTimestamp[21] := BenchUut2.FaultTimestamp;
   TraceIn_CycleTime[21] := BenchUut2.CycleTime;
   BenchUut2();
   TraceOut_THICKNESS_ALARM[21] := BenchUut2.THICKNESS_ALARM;
   TraceOut_Slab_Fault_Counter[21] := BenchUut2.Slab_Fault_Counter;
   TraceOut_Slab_Runtime_Accumulator[21] := BenchUut2.Slab_Runtime_Accumulator;
   TraceOut_Slab_Fault_History_0[21] := BenchUut2.Slab_Fault_History[0];
   TraceOut_Slab_Fault_History_1[21] := BenchUut2.Slab_Fault_History[1];
   TraceOut_Slab_Fault_History_2[21] := BenchUut2.Slab_Fault_History[2];
   TraceOut_Slab_Fault_History_3[21] := BenchUut2.Slab_Fault_History[3];
   TraceOut_Slab_Fault_History_4[21] := BenchUut2.Slab_Fault_History[4];
   BenchCalls := BenchCalls + 1;
   BenchStep := BenchStep + 1;
  END_IF;
 22:
  IF BenchCurrentTime - BenchLastTime >= UDINT_TO_TIME(100) THEN
   TraceDt[22] := TIME_TO_UDINT(BenchCurrentTime - BenchLastTime);
   BenchLastTime := BenchCurrentTime;
   BenchUut2.THICKNESS_FAULT := TRUE;
   BenchUut2.THICKNESS_SIGNAL_VALID := TRUE;
   BenchUut2.CUTTING_RUN := TRUE;
   BenchUut2.FaultTimestamp := DINT#0;
   BenchUut2.CycleTime := T#100ms;
   TraceIn_THICKNESS_FAULT[22] := BenchUut2.THICKNESS_FAULT;
   TraceIn_THICKNESS_SIGNAL_VALID[22] := BenchUut2.THICKNESS_SIGNAL_VALID;
   TraceIn_CUTTING_RUN[22] := BenchUut2.CUTTING_RUN;
   TraceIn_FaultTimestamp[22] := BenchUut2.FaultTimestamp;
   TraceIn_CycleTime[22] := BenchUut2.CycleTime;
   BenchUut2();
   TraceOut_THICKNESS_ALARM[22] := BenchUut2.THICKNESS_ALARM;
   TraceOut_Slab_Fault_Counter[22] := BenchUut2.Slab_Fault_Counter;
   TraceOut_Slab_Runtime_Accumulator[22] := BenchUut2.Slab_Runtime_Accumulator;
   TraceOut_Slab_Fault_History_0[22] := BenchUut2.Slab_Fault_History[0];
   TraceOut_Slab_Fault_History_1[22] := BenchUut2.Slab_Fault_History[1];
   TraceOut_Slab_Fault_History_2[22] := BenchUut2.Slab_Fault_History[2];
   TraceOut_Slab_Fault_History_3[22] := BenchUut2.Slab_Fault_History[3];
   TraceOut_Slab_Fault_History_4[22] := BenchUut2.Slab_Fault_History[4];
   BenchCalls := BenchCalls + 1;
   BenchStep := BenchStep + 1;
  END_IF;
 23:
  IF BenchCurrentTime - BenchLastTime >= UDINT_TO_TIME(100) THEN
   TraceDt[23] := TIME_TO_UDINT(BenchCurrentTime - BenchLastTime);
   BenchLastTime := BenchCurrentTime;
   BenchUut2.THICKNESS_FAULT := FALSE;
   BenchUut2.THICKNESS_SIGNAL_VALID := FALSE;
   BenchUut2.CUTTING_RUN := TRUE;
   BenchUut2.FaultTimestamp := DINT#0;
   BenchUut2.CycleTime := T#100ms;
   TraceIn_THICKNESS_FAULT[23] := BenchUut2.THICKNESS_FAULT;
   TraceIn_THICKNESS_SIGNAL_VALID[23] := BenchUut2.THICKNESS_SIGNAL_VALID;
   TraceIn_CUTTING_RUN[23] := BenchUut2.CUTTING_RUN;
   TraceIn_FaultTimestamp[23] := BenchUut2.FaultTimestamp;
   TraceIn_CycleTime[23] := BenchUut2.CycleTime;
   BenchUut2();
   TraceOut_THICKNESS_ALARM[23] := BenchUut2.THICKNESS_ALARM;
   TraceOut_Slab_Fault_Counter[23] := BenchUut2.Slab_Fault_Counter;
   TraceOut_Slab_Runtime_Accumulator[23] := BenchUut2.Slab_Runtime_Accumulator;
   TraceOut_Slab_Fault_History_0[23] := BenchUut2.Slab_Fault_History[0];
   TraceOut_Slab_Fault_History_1[23] := BenchUut2.Slab_Fault_History[1];
   TraceOut_Slab_Fault_History_2[23] := BenchUut2.Slab_Fault_History[2];
   TraceOut_Slab_Fault_History_3[23] := BenchUut2.Slab_Fault_History[3];
   TraceOut_Slab_Fault_History_4[23] := BenchUut2.Slab_Fault_History[4];
   BenchCalls := BenchCalls + 1;
   BenchStep := BenchStep + 1;
  END_IF;
 24:
  IF BenchCurrentTime - BenchLastTime >= UDINT_TO_TIME(100) THEN
   TraceDt[24] := TIME_TO_UDINT(BenchCurrentTime - BenchLastTime);
   BenchLastTime := BenchCurrentTime;
   BenchUut2.THICKNESS_FAULT := FALSE;
   BenchUut2.THICKNESS_SIGNAL_VALID := TRUE;
   BenchUut2.CUTTING_RUN := FALSE;
   BenchUut2.FaultTimestamp := DINT#0;
   BenchUut2.CycleTime := T#100ms;
   TraceIn_THICKNESS_FAULT[24] := BenchUut2.THICKNESS_FAULT;
   TraceIn_THICKNESS_SIGNAL_VALID[24] := BenchUut2.THICKNESS_SIGNAL_VALID;
   TraceIn_CUTTING_RUN[24] := BenchUut2.CUTTING_RUN;
   TraceIn_FaultTimestamp[24] := BenchUut2.FaultTimestamp;
   TraceIn_CycleTime[24] := BenchUut2.CycleTime;
   BenchUut2();
   TraceOut_THICKNESS_ALARM[24] := BenchUut2.THICKNESS_ALARM;
   TraceOut_Slab_Fault_Counter[24] := BenchUut2.Slab_Fault_Counter;
   TraceOut_Slab_Runtime_Accumulator[24] := BenchUut2.Slab_Runtime_Accumulator;
   TraceOut_Slab_Fault_History_0[24] := BenchUut2.Slab_Fault_History[0];
   TraceOut_Slab_Fault_History_1[24] := BenchUut2.Slab_Fault_History[1];
   TraceOut_Slab_Fault_History_2[24] := BenchUut2.Slab_Fault_History[2];
   TraceOut_Slab_Fault_History_3[24] := BenchUut2.Slab_Fault_History[3];
   TraceOut_Slab_Fault_History_4[24] := BenchUut2.Slab_Fault_History[4];
   BenchCalls := BenchCalls + 1;
   BenchStep := BenchStep + 1;
  END_IF;
 25:
  IF BenchCurrentTime - BenchLastTime >= UDINT_TO_TIME(0) THEN
   TraceDt[25] := TIME_TO_UDINT(BenchCurrentTime - BenchLastTime);
   BenchLastTime := BenchCurrentTime;
   BenchUut3.THICKNESS_FAULT := TRUE;
   BenchUut3.THICKNESS_SIGNAL_VALID := TRUE;
   BenchUut3.CUTTING_RUN := TRUE;
   BenchUut3.FaultTimestamp := DINT#10;
   BenchUut3.CycleTime := T#100ms;
   TraceIn_THICKNESS_FAULT[25] := BenchUut3.THICKNESS_FAULT;
   TraceIn_THICKNESS_SIGNAL_VALID[25] := BenchUut3.THICKNESS_SIGNAL_VALID;
   TraceIn_CUTTING_RUN[25] := BenchUut3.CUTTING_RUN;
   TraceIn_FaultTimestamp[25] := BenchUut3.FaultTimestamp;
   TraceIn_CycleTime[25] := BenchUut3.CycleTime;
   BenchUut3();
   TraceOut_THICKNESS_ALARM[25] := BenchUut3.THICKNESS_ALARM;
   TraceOut_Slab_Fault_Counter[25] := BenchUut3.Slab_Fault_Counter;
   TraceOut_Slab_Runtime_Accumulator[25] := BenchUut3.Slab_Runtime_Accumulator;
   TraceOut_Slab_Fault_History_0[25] := BenchUut3.Slab_Fault_History[0];
   TraceOut_Slab_Fault_History_1[25] := BenchUut3.Slab_Fault_History[1];
   TraceOut_Slab_Fault_History_2[25] := BenchUut3.Slab_Fault_History[2];
   TraceOut_Slab_Fault_History_3[25] := BenchUut3.Slab_Fault_History[3];
   TraceOut_Slab_Fault_History_4[25] := BenchUut3.Slab_Fault_History[4];
   BenchCalls := BenchCalls + 1;
   BenchStep := BenchStep + 1;
  END_IF;
 26:
  IF BenchCurrentTime - BenchLastTime >= UDINT_TO_TIME(400) THEN
   TraceDt[26] := TIME_TO_UDINT(BenchCurrentTime - BenchLastTime);
   BenchLastTime := BenchCurrentTime;
   BenchUut3.THICKNESS_FAULT := FALSE;
   BenchUut3.THICKNESS_SIGNAL_VALID := TRUE;
   BenchUut3.CUTTING_RUN := TRUE;
   BenchUut3.FaultTimestamp := DINT#10;
   BenchUut3.CycleTime := T#400ms;
   TraceIn_THICKNESS_FAULT[26] := BenchUut3.THICKNESS_FAULT;
   TraceIn_THICKNESS_SIGNAL_VALID[26] := BenchUut3.THICKNESS_SIGNAL_VALID;
   TraceIn_CUTTING_RUN[26] := BenchUut3.CUTTING_RUN;
   TraceIn_FaultTimestamp[26] := BenchUut3.FaultTimestamp;
   TraceIn_CycleTime[26] := BenchUut3.CycleTime;
   BenchUut3();
   TraceOut_THICKNESS_ALARM[26] := BenchUut3.THICKNESS_ALARM;
   TraceOut_Slab_Fault_Counter[26] := BenchUut3.Slab_Fault_Counter;
   TraceOut_Slab_Runtime_Accumulator[26] := BenchUut3.Slab_Runtime_Accumulator;
   TraceOut_Slab_Fault_History_0[26] := BenchUut3.Slab_Fault_History[0];
   TraceOut_Slab_Fault_History_1[26] := BenchUut3.Slab_Fault_History[1];
   TraceOut_Slab_Fault_History_2[26] := BenchUut3.Slab_Fault_History[2];
   TraceOut_Slab_Fault_History_3[26] := BenchUut3.Slab_Fault_History[3];
   TraceOut_Slab_Fault_History_4[26] := BenchUut3.Slab_Fault_History[4];
   BenchCalls := BenchCalls + 1;
   BenchStep := BenchStep + 1;
  END_IF;
 27:
  IF BenchCurrentTime - BenchLastTime >= UDINT_TO_TIME(50) THEN
   TraceDt[27] := TIME_TO_UDINT(BenchCurrentTime - BenchLastTime);
   BenchLastTime := BenchCurrentTime;
   BenchUut3.THICKNESS_FAULT := TRUE;
   BenchUut3.THICKNESS_SIGNAL_VALID := TRUE;
   BenchUut3.CUTTING_RUN := TRUE;
   BenchUut3.FaultTimestamp := DINT#20;
   BenchUut3.CycleTime := T#50ms;
   TraceIn_THICKNESS_FAULT[27] := BenchUut3.THICKNESS_FAULT;
   TraceIn_THICKNESS_SIGNAL_VALID[27] := BenchUut3.THICKNESS_SIGNAL_VALID;
   TraceIn_CUTTING_RUN[27] := BenchUut3.CUTTING_RUN;
   TraceIn_FaultTimestamp[27] := BenchUut3.FaultTimestamp;
   TraceIn_CycleTime[27] := BenchUut3.CycleTime;
   BenchUut3();
   TraceOut_THICKNESS_ALARM[27] := BenchUut3.THICKNESS_ALARM;
   TraceOut_Slab_Fault_Counter[27] := BenchUut3.Slab_Fault_Counter;
   TraceOut_Slab_Runtime_Accumulator[27] := BenchUut3.Slab_Runtime_Accumulator;
   TraceOut_Slab_Fault_History_0[27] := BenchUut3.Slab_Fault_History[0];
   TraceOut_Slab_Fault_History_1[27] := BenchUut3.Slab_Fault_History[1];
   TraceOut_Slab_Fault_History_2[27] := BenchUut3.Slab_Fault_History[2];
   TraceOut_Slab_Fault_History_3[27] := BenchUut3.Slab_Fault_History[3];
   TraceOut_Slab_Fault_History_4[27] := BenchUut3.Slab_Fault_History[4];
   BenchCalls := BenchCalls + 1;
   BenchStep := BenchStep + 1;
  END_IF;
 28:
  IF BenchCurrentTime - BenchLastTime >= UDINT_TO_TIME(499) THEN
   TraceDt[28] := TIME_TO_UDINT(BenchCurrentTime - BenchLastTime);
   BenchLastTime := BenchCurrentTime;
   BenchUut3.THICKNESS_FAULT := FALSE;
   BenchUut3.THICKNESS_SIGNAL_VALID := TRUE;
   BenchUut3.CUTTING_RUN := TRUE;
   BenchUut3.FaultTimestamp := DINT#20;
   BenchUut3.CycleTime := T#499ms;
   TraceIn_THICKNESS_FAULT[28] := BenchUut3.THICKNESS_FAULT;
   TraceIn_THICKNESS_SIGNAL_VALID[28] := BenchUut3.THICKNESS_SIGNAL_VALID;
   TraceIn_CUTTING_RUN[28] := BenchUut3.CUTTING_RUN;
   TraceIn_FaultTimestamp[28] := BenchUut3.FaultTimestamp;
   TraceIn_CycleTime[28] := BenchUut3.CycleTime;
   BenchUut3();
   TraceOut_THICKNESS_ALARM[28] := BenchUut3.THICKNESS_ALARM;
   TraceOut_Slab_Fault_Counter[28] := BenchUut3.Slab_Fault_Counter;
   TraceOut_Slab_Runtime_Accumulator[28] := BenchUut3.Slab_Runtime_Accumulator;
   TraceOut_Slab_Fault_History_0[28] := BenchUut3.Slab_Fault_History[0];
   TraceOut_Slab_Fault_History_1[28] := BenchUut3.Slab_Fault_History[1];
   TraceOut_Slab_Fault_History_2[28] := BenchUut3.Slab_Fault_History[2];
   TraceOut_Slab_Fault_History_3[28] := BenchUut3.Slab_Fault_History[3];
   TraceOut_Slab_Fault_History_4[28] := BenchUut3.Slab_Fault_History[4];
   BenchCalls := BenchCalls + 1;
   BenchStep := BenchStep + 1;
  END_IF;
 29:
  IF BenchCurrentTime - BenchLastTime >= UDINT_TO_TIME(1) THEN
   TraceDt[29] := TIME_TO_UDINT(BenchCurrentTime - BenchLastTime);
   BenchLastTime := BenchCurrentTime;
   BenchUut3.THICKNESS_FAULT := FALSE;
   BenchUut3.THICKNESS_SIGNAL_VALID := TRUE;
   BenchUut3.CUTTING_RUN := TRUE;
   BenchUut3.FaultTimestamp := DINT#20;
   BenchUut3.CycleTime := T#1ms;
   TraceIn_THICKNESS_FAULT[29] := BenchUut3.THICKNESS_FAULT;
   TraceIn_THICKNESS_SIGNAL_VALID[29] := BenchUut3.THICKNESS_SIGNAL_VALID;
   TraceIn_CUTTING_RUN[29] := BenchUut3.CUTTING_RUN;
   TraceIn_FaultTimestamp[29] := BenchUut3.FaultTimestamp;
   TraceIn_CycleTime[29] := BenchUut3.CycleTime;
   BenchUut3();
   TraceOut_THICKNESS_ALARM[29] := BenchUut3.THICKNESS_ALARM;
   TraceOut_Slab_Fault_Counter[29] := BenchUut3.Slab_Fault_Counter;
   TraceOut_Slab_Runtime_Accumulator[29] := BenchUut3.Slab_Runtime_Accumulator;
   TraceOut_Slab_Fault_History_0[29] := BenchUut3.Slab_Fault_History[0];
   TraceOut_Slab_Fault_History_1[29] := BenchUut3.Slab_Fault_History[1];
   TraceOut_Slab_Fault_History_2[29] := BenchUut3.Slab_Fault_History[2];
   TraceOut_Slab_Fault_History_3[29] := BenchUut3.Slab_Fault_History[3];
   TraceOut_Slab_Fault_History_4[29] := BenchUut3.Slab_Fault_History[4];
   BenchCalls := BenchCalls + 1;
   BenchStep := BenchStep + 1;
  END_IF;
 30:
  IF BenchCurrentTime - BenchLastTime >= UDINT_TO_TIME(100) THEN
   TraceDt[30] := TIME_TO_UDINT(BenchCurrentTime - BenchLastTime);
   BenchLastTime := BenchCurrentTime;
   BenchUut3.THICKNESS_FAULT := TRUE;
   BenchUut3.THICKNESS_SIGNAL_VALID := TRUE;
   BenchUut3.CUTTING_RUN := FALSE;
   BenchUut3.FaultTimestamp := DINT#30;
   BenchUut3.CycleTime := T#100ms;
   TraceIn_THICKNESS_FAULT[30] := BenchUut3.THICKNESS_FAULT;
   TraceIn_THICKNESS_SIGNAL_VALID[30] := BenchUut3.THICKNESS_SIGNAL_VALID;
   TraceIn_CUTTING_RUN[30] := BenchUut3.CUTTING_RUN;
   TraceIn_FaultTimestamp[30] := BenchUut3.FaultTimestamp;
   TraceIn_CycleTime[30] := BenchUut3.CycleTime;
   BenchUut3();
   TraceOut_THICKNESS_ALARM[30] := BenchUut3.THICKNESS_ALARM;
   TraceOut_Slab_Fault_Counter[30] := BenchUut3.Slab_Fault_Counter;
   TraceOut_Slab_Runtime_Accumulator[30] := BenchUut3.Slab_Runtime_Accumulator;
   TraceOut_Slab_Fault_History_0[30] := BenchUut3.Slab_Fault_History[0];
   TraceOut_Slab_Fault_History_1[30] := BenchUut3.Slab_Fault_History[1];
   TraceOut_Slab_Fault_History_2[30] := BenchUut3.Slab_Fault_History[2];
   TraceOut_Slab_Fault_History_3[30] := BenchUut3.Slab_Fault_History[3];
   TraceOut_Slab_Fault_History_4[30] := BenchUut3.Slab_Fault_History[4];
   BenchCalls := BenchCalls + 1;
   BenchStep := BenchStep + 1;
  END_IF;
 31:
  IF BenchCurrentTime - BenchLastTime >= UDINT_TO_TIME(600) THEN
   TraceDt[31] := TIME_TO_UDINT(BenchCurrentTime - BenchLastTime);
   BenchLastTime := BenchCurrentTime;
   BenchUut3.THICKNESS_FAULT := TRUE;
   BenchUut3.THICKNESS_SIGNAL_VALID := TRUE;
   BenchUut3.CUTTING_RUN := FALSE;
   BenchUut3.FaultTimestamp := DINT#30;
   BenchUut3.CycleTime := T#600ms;
   TraceIn_THICKNESS_FAULT[31] := BenchUut3.THICKNESS_FAULT;
   TraceIn_THICKNESS_SIGNAL_VALID[31] := BenchUut3.THICKNESS_SIGNAL_VALID;
   TraceIn_CUTTING_RUN[31] := BenchUut3.CUTTING_RUN;
   TraceIn_FaultTimestamp[31] := BenchUut3.FaultTimestamp;
   TraceIn_CycleTime[31] := BenchUut3.CycleTime;
   BenchUut3();
   TraceOut_THICKNESS_ALARM[31] := BenchUut3.THICKNESS_ALARM;
   TraceOut_Slab_Fault_Counter[31] := BenchUut3.Slab_Fault_Counter;
   TraceOut_Slab_Runtime_Accumulator[31] := BenchUut3.Slab_Runtime_Accumulator;
   TraceOut_Slab_Fault_History_0[31] := BenchUut3.Slab_Fault_History[0];
   TraceOut_Slab_Fault_History_1[31] := BenchUut3.Slab_Fault_History[1];
   TraceOut_Slab_Fault_History_2[31] := BenchUut3.Slab_Fault_History[2];
   TraceOut_Slab_Fault_History_3[31] := BenchUut3.Slab_Fault_History[3];
   TraceOut_Slab_Fault_History_4[31] := BenchUut3.Slab_Fault_History[4];
   BenchCalls := BenchCalls + 1;
   BenchStep := BenchStep + 1;
  END_IF;
 32:
  IF BenchCurrentTime - BenchLastTime >= UDINT_TO_TIME(10) THEN
   TraceDt[32] := TIME_TO_UDINT(BenchCurrentTime - BenchLastTime);
   BenchLastTime := BenchCurrentTime;
   BenchUut3.THICKNESS_FAULT := FALSE;
   BenchUut3.THICKNESS_SIGNAL_VALID := TRUE;
   BenchUut3.CUTTING_RUN := TRUE;
   BenchUut3.FaultTimestamp := DINT#30;
   BenchUut3.CycleTime := T#10ms;
   TraceIn_THICKNESS_FAULT[32] := BenchUut3.THICKNESS_FAULT;
   TraceIn_THICKNESS_SIGNAL_VALID[32] := BenchUut3.THICKNESS_SIGNAL_VALID;
   TraceIn_CUTTING_RUN[32] := BenchUut3.CUTTING_RUN;
   TraceIn_FaultTimestamp[32] := BenchUut3.FaultTimestamp;
   TraceIn_CycleTime[32] := BenchUut3.CycleTime;
   BenchUut3();
   TraceOut_THICKNESS_ALARM[32] := BenchUut3.THICKNESS_ALARM;
   TraceOut_Slab_Fault_Counter[32] := BenchUut3.Slab_Fault_Counter;
   TraceOut_Slab_Runtime_Accumulator[32] := BenchUut3.Slab_Runtime_Accumulator;
   TraceOut_Slab_Fault_History_0[32] := BenchUut3.Slab_Fault_History[0];
   TraceOut_Slab_Fault_History_1[32] := BenchUut3.Slab_Fault_History[1];
   TraceOut_Slab_Fault_History_2[32] := BenchUut3.Slab_Fault_History[2];
   TraceOut_Slab_Fault_History_3[32] := BenchUut3.Slab_Fault_History[3];
   TraceOut_Slab_Fault_History_4[32] := BenchUut3.Slab_Fault_History[4];
   BenchCalls := BenchCalls + 1;
   BenchStep := BenchStep + 1;
  END_IF;
 33:
  IF BenchCurrentTime - BenchLastTime >= UDINT_TO_TIME(50) THEN
   TraceDt[33] := TIME_TO_UDINT(BenchCurrentTime - BenchLastTime);
   BenchLastTime := BenchCurrentTime;
   BenchUut3.THICKNESS_FAULT := TRUE;
   BenchUut3.THICKNESS_SIGNAL_VALID := TRUE;
   BenchUut3.CUTTING_RUN := FALSE;
   BenchUut3.FaultTimestamp := DINT#40;
   BenchUut3.CycleTime := T#50ms;
   TraceIn_THICKNESS_FAULT[33] := BenchUut3.THICKNESS_FAULT;
   TraceIn_THICKNESS_SIGNAL_VALID[33] := BenchUut3.THICKNESS_SIGNAL_VALID;
   TraceIn_CUTTING_RUN[33] := BenchUut3.CUTTING_RUN;
   TraceIn_FaultTimestamp[33] := BenchUut3.FaultTimestamp;
   TraceIn_CycleTime[33] := BenchUut3.CycleTime;
   BenchUut3();
   TraceOut_THICKNESS_ALARM[33] := BenchUut3.THICKNESS_ALARM;
   TraceOut_Slab_Fault_Counter[33] := BenchUut3.Slab_Fault_Counter;
   TraceOut_Slab_Runtime_Accumulator[33] := BenchUut3.Slab_Runtime_Accumulator;
   TraceOut_Slab_Fault_History_0[33] := BenchUut3.Slab_Fault_History[0];
   TraceOut_Slab_Fault_History_1[33] := BenchUut3.Slab_Fault_History[1];
   TraceOut_Slab_Fault_History_2[33] := BenchUut3.Slab_Fault_History[2];
   TraceOut_Slab_Fault_History_3[33] := BenchUut3.Slab_Fault_History[3];
   TraceOut_Slab_Fault_History_4[33] := BenchUut3.Slab_Fault_History[4];
   BenchCalls := BenchCalls + 1;
   BenchStep := BenchStep + 1;
  END_IF;
 34:
  IF BenchCurrentTime - BenchLastTime >= UDINT_TO_TIME(50) THEN
   TraceDt[34] := TIME_TO_UDINT(BenchCurrentTime - BenchLastTime);
   BenchLastTime := BenchCurrentTime;
   BenchUut3.THICKNESS_FAULT := FALSE;
   BenchUut3.THICKNESS_SIGNAL_VALID := FALSE;
   BenchUut3.CUTTING_RUN := TRUE;
   BenchUut3.FaultTimestamp := DINT#40;
   BenchUut3.CycleTime := T#50ms;
   TraceIn_THICKNESS_FAULT[34] := BenchUut3.THICKNESS_FAULT;
   TraceIn_THICKNESS_SIGNAL_VALID[34] := BenchUut3.THICKNESS_SIGNAL_VALID;
   TraceIn_CUTTING_RUN[34] := BenchUut3.CUTTING_RUN;
   TraceIn_FaultTimestamp[34] := BenchUut3.FaultTimestamp;
   TraceIn_CycleTime[34] := BenchUut3.CycleTime;
   BenchUut3();
   TraceOut_THICKNESS_ALARM[34] := BenchUut3.THICKNESS_ALARM;
   TraceOut_Slab_Fault_Counter[34] := BenchUut3.Slab_Fault_Counter;
   TraceOut_Slab_Runtime_Accumulator[34] := BenchUut3.Slab_Runtime_Accumulator;
   TraceOut_Slab_Fault_History_0[34] := BenchUut3.Slab_Fault_History[0];
   TraceOut_Slab_Fault_History_1[34] := BenchUut3.Slab_Fault_History[1];
   TraceOut_Slab_Fault_History_2[34] := BenchUut3.Slab_Fault_History[2];
   TraceOut_Slab_Fault_History_3[34] := BenchUut3.Slab_Fault_History[3];
   TraceOut_Slab_Fault_History_4[34] := BenchUut3.Slab_Fault_History[4];
   BenchCalls := BenchCalls + 1;
   BenchStep := BenchStep + 1;
  END_IF;
 35:
  IF BenchCurrentTime - BenchLastTime >= UDINT_TO_TIME(50) THEN
   TraceDt[35] := TIME_TO_UDINT(BenchCurrentTime - BenchLastTime);
   BenchLastTime := BenchCurrentTime;
   BenchUut3.THICKNESS_FAULT := FALSE;
   BenchUut3.THICKNESS_SIGNAL_VALID := TRUE;
   BenchUut3.CUTTING_RUN := TRUE;
   BenchUut3.FaultTimestamp := DINT#40;
   BenchUut3.CycleTime := T#50ms;
   TraceIn_THICKNESS_FAULT[35] := BenchUut3.THICKNESS_FAULT;
   TraceIn_THICKNESS_SIGNAL_VALID[35] := BenchUut3.THICKNESS_SIGNAL_VALID;
   TraceIn_CUTTING_RUN[35] := BenchUut3.CUTTING_RUN;
   TraceIn_FaultTimestamp[35] := BenchUut3.FaultTimestamp;
   TraceIn_CycleTime[35] := BenchUut3.CycleTime;
   BenchUut3();
   TraceOut_THICKNESS_ALARM[35] := BenchUut3.THICKNESS_ALARM;
   TraceOut_Slab_Fault_Counter[35] := BenchUut3.Slab_Fault_Counter;
   TraceOut_Slab_Runtime_Accumulator[35] := BenchUut3.Slab_Runtime_Accumulator;
   TraceOut_Slab_Fault_History_0[35] := BenchUut3.Slab_Fault_History[0];
   TraceOut_Slab_Fault_History_1[35] := BenchUut3.Slab_Fault_History[1];
   TraceOut_Slab_Fault_History_2[35] := BenchUut3.Slab_Fault_History[2];
   TraceOut_Slab_Fault_History_3[35] := BenchUut3.Slab_Fault_History[3];
   TraceOut_Slab_Fault_History_4[35] := BenchUut3.Slab_Fault_History[4];
   BenchCalls := BenchCalls + 1;
   BenchStep := BenchStep + 1;
  END_IF;
 36:
  IF BenchCurrentTime - BenchLastTime >= UDINT_TO_TIME(0) THEN
   TraceDt[36] := TIME_TO_UDINT(BenchCurrentTime - BenchLastTime);
   BenchLastTime := BenchCurrentTime;
   BenchUut4.THICKNESS_FAULT := TRUE;
   BenchUut4.THICKNESS_SIGNAL_VALID := TRUE;
   BenchUut4.CUTTING_RUN := FALSE;
   BenchUut4.FaultTimestamp := DINT#10;
   BenchUut4.CycleTime := T#100ms;
   TraceIn_THICKNESS_FAULT[36] := BenchUut4.THICKNESS_FAULT;
   TraceIn_THICKNESS_SIGNAL_VALID[36] := BenchUut4.THICKNESS_SIGNAL_VALID;
   TraceIn_CUTTING_RUN[36] := BenchUut4.CUTTING_RUN;
   TraceIn_FaultTimestamp[36] := BenchUut4.FaultTimestamp;
   TraceIn_CycleTime[36] := BenchUut4.CycleTime;
   BenchUut4();
   TraceOut_THICKNESS_ALARM[36] := BenchUut4.THICKNESS_ALARM;
   TraceOut_Slab_Fault_Counter[36] := BenchUut4.Slab_Fault_Counter;
   TraceOut_Slab_Runtime_Accumulator[36] := BenchUut4.Slab_Runtime_Accumulator;
   TraceOut_Slab_Fault_History_0[36] := BenchUut4.Slab_Fault_History[0];
   TraceOut_Slab_Fault_History_1[36] := BenchUut4.Slab_Fault_History[1];
   TraceOut_Slab_Fault_History_2[36] := BenchUut4.Slab_Fault_History[2];
   TraceOut_Slab_Fault_History_3[36] := BenchUut4.Slab_Fault_History[3];
   TraceOut_Slab_Fault_History_4[36] := BenchUut4.Slab_Fault_History[4];
   BenchCalls := BenchCalls + 1;
   BenchStep := BenchStep + 1;
  END_IF;
 37:
  IF BenchCurrentTime - BenchLastTime >= UDINT_TO_TIME(100) THEN
   TraceDt[37] := TIME_TO_UDINT(BenchCurrentTime - BenchLastTime);
   BenchLastTime := BenchCurrentTime;
   BenchUut4.THICKNESS_FAULT := TRUE;
   BenchUut4.THICKNESS_SIGNAL_VALID := TRUE;
   BenchUut4.CUTTING_RUN := FALSE;
   BenchUut4.FaultTimestamp := DINT#10;
   BenchUut4.CycleTime := T#100ms;
   TraceIn_THICKNESS_FAULT[37] := BenchUut4.THICKNESS_FAULT;
   TraceIn_THICKNESS_SIGNAL_VALID[37] := BenchUut4.THICKNESS_SIGNAL_VALID;
   TraceIn_CUTTING_RUN[37] := BenchUut4.CUTTING_RUN;
   TraceIn_FaultTimestamp[37] := BenchUut4.FaultTimestamp;
   TraceIn_CycleTime[37] := BenchUut4.CycleTime;
   BenchUut4();
   TraceOut_THICKNESS_ALARM[37] := BenchUut4.THICKNESS_ALARM;
   TraceOut_Slab_Fault_Counter[37] := BenchUut4.Slab_Fault_Counter;
   TraceOut_Slab_Runtime_Accumulator[37] := BenchUut4.Slab_Runtime_Accumulator;
   TraceOut_Slab_Fault_History_0[37] := BenchUut4.Slab_Fault_History[0];
   TraceOut_Slab_Fault_History_1[37] := BenchUut4.Slab_Fault_History[1];
   TraceOut_Slab_Fault_History_2[37] := BenchUut4.Slab_Fault_History[2];
   TraceOut_Slab_Fault_History_3[37] := BenchUut4.Slab_Fault_History[3];
   TraceOut_Slab_Fault_History_4[37] := BenchUut4.Slab_Fault_History[4];
   BenchCalls := BenchCalls + 1;
   BenchStep := BenchStep + 1;
  END_IF;
 38:
  IF BenchCurrentTime - BenchLastTime >= UDINT_TO_TIME(100) THEN
   TraceDt[38] := TIME_TO_UDINT(BenchCurrentTime - BenchLastTime);
   BenchLastTime := BenchCurrentTime;
   BenchUut4.THICKNESS_FAULT := TRUE;
   BenchUut4.THICKNESS_SIGNAL_VALID := TRUE;
   BenchUut4.CUTTING_RUN := FALSE;
   BenchUut4.FaultTimestamp := DINT#10;
   BenchUut4.CycleTime := T#100ms;
   TraceIn_THICKNESS_FAULT[38] := BenchUut4.THICKNESS_FAULT;
   TraceIn_THICKNESS_SIGNAL_VALID[38] := BenchUut4.THICKNESS_SIGNAL_VALID;
   TraceIn_CUTTING_RUN[38] := BenchUut4.CUTTING_RUN;
   TraceIn_FaultTimestamp[38] := BenchUut4.FaultTimestamp;
   TraceIn_CycleTime[38] := BenchUut4.CycleTime;
   BenchUut4();
   TraceOut_THICKNESS_ALARM[38] := BenchUut4.THICKNESS_ALARM;
   TraceOut_Slab_Fault_Counter[38] := BenchUut4.Slab_Fault_Counter;
   TraceOut_Slab_Runtime_Accumulator[38] := BenchUut4.Slab_Runtime_Accumulator;
   TraceOut_Slab_Fault_History_0[38] := BenchUut4.Slab_Fault_History[0];
   TraceOut_Slab_Fault_History_1[38] := BenchUut4.Slab_Fault_History[1];
   TraceOut_Slab_Fault_History_2[38] := BenchUut4.Slab_Fault_History[2];
   TraceOut_Slab_Fault_History_3[38] := BenchUut4.Slab_Fault_History[3];
   TraceOut_Slab_Fault_History_4[38] := BenchUut4.Slab_Fault_History[4];
   BenchCalls := BenchCalls + 1;
   BenchStep := BenchStep + 1;
  END_IF;
 39:
  IF BenchCurrentTime - BenchLastTime >= UDINT_TO_TIME(100) THEN
   TraceDt[39] := TIME_TO_UDINT(BenchCurrentTime - BenchLastTime);
   BenchLastTime := BenchCurrentTime;
   BenchUut4.THICKNESS_FAULT := FALSE;
   BenchUut4.THICKNESS_SIGNAL_VALID := TRUE;
   BenchUut4.CUTTING_RUN := FALSE;
   BenchUut4.FaultTimestamp := DINT#10;
   BenchUut4.CycleTime := T#100ms;
   TraceIn_THICKNESS_FAULT[39] := BenchUut4.THICKNESS_FAULT;
   TraceIn_THICKNESS_SIGNAL_VALID[39] := BenchUut4.THICKNESS_SIGNAL_VALID;
   TraceIn_CUTTING_RUN[39] := BenchUut4.CUTTING_RUN;
   TraceIn_FaultTimestamp[39] := BenchUut4.FaultTimestamp;
   TraceIn_CycleTime[39] := BenchUut4.CycleTime;
   BenchUut4();
   TraceOut_THICKNESS_ALARM[39] := BenchUut4.THICKNESS_ALARM;
   TraceOut_Slab_Fault_Counter[39] := BenchUut4.Slab_Fault_Counter;
   TraceOut_Slab_Runtime_Accumulator[39] := BenchUut4.Slab_Runtime_Accumulator;
   TraceOut_Slab_Fault_History_0[39] := BenchUut4.Slab_Fault_History[0];
   TraceOut_Slab_Fault_History_1[39] := BenchUut4.Slab_Fault_History[1];
   TraceOut_Slab_Fault_History_2[39] := BenchUut4.Slab_Fault_History[2];
   TraceOut_Slab_Fault_History_3[39] := BenchUut4.Slab_Fault_History[3];
   TraceOut_Slab_Fault_History_4[39] := BenchUut4.Slab_Fault_History[4];
   BenchCalls := BenchCalls + 1;
   BenchStep := BenchStep + 1;
  END_IF;
 40:
  IF BenchCurrentTime - BenchLastTime >= UDINT_TO_TIME(100) THEN
   TraceDt[40] := TIME_TO_UDINT(BenchCurrentTime - BenchLastTime);
   BenchLastTime := BenchCurrentTime;
   BenchUut4.THICKNESS_FAULT := TRUE;
   BenchUut4.THICKNESS_SIGNAL_VALID := TRUE;
   BenchUut4.CUTTING_RUN := FALSE;
   BenchUut4.FaultTimestamp := DINT#20;
   BenchUut4.CycleTime := T#100ms;
   TraceIn_THICKNESS_FAULT[40] := BenchUut4.THICKNESS_FAULT;
   TraceIn_THICKNESS_SIGNAL_VALID[40] := BenchUut4.THICKNESS_SIGNAL_VALID;
   TraceIn_CUTTING_RUN[40] := BenchUut4.CUTTING_RUN;
   TraceIn_FaultTimestamp[40] := BenchUut4.FaultTimestamp;
   TraceIn_CycleTime[40] := BenchUut4.CycleTime;
   BenchUut4();
   TraceOut_THICKNESS_ALARM[40] := BenchUut4.THICKNESS_ALARM;
   TraceOut_Slab_Fault_Counter[40] := BenchUut4.Slab_Fault_Counter;
   TraceOut_Slab_Runtime_Accumulator[40] := BenchUut4.Slab_Runtime_Accumulator;
   TraceOut_Slab_Fault_History_0[40] := BenchUut4.Slab_Fault_History[0];
   TraceOut_Slab_Fault_History_1[40] := BenchUut4.Slab_Fault_History[1];
   TraceOut_Slab_Fault_History_2[40] := BenchUut4.Slab_Fault_History[2];
   TraceOut_Slab_Fault_History_3[40] := BenchUut4.Slab_Fault_History[3];
   TraceOut_Slab_Fault_History_4[40] := BenchUut4.Slab_Fault_History[4];
   BenchCalls := BenchCalls + 1;
   BenchStep := BenchStep + 1;
  END_IF;
 41:
  IF BenchCurrentTime - BenchLastTime >= UDINT_TO_TIME(100) THEN
   TraceDt[41] := TIME_TO_UDINT(BenchCurrentTime - BenchLastTime);
   BenchLastTime := BenchCurrentTime;
   BenchUut4.THICKNESS_FAULT := FALSE;
   BenchUut4.THICKNESS_SIGNAL_VALID := TRUE;
   BenchUut4.CUTTING_RUN := FALSE;
   BenchUut4.FaultTimestamp := DINT#20;
   BenchUut4.CycleTime := T#100ms;
   TraceIn_THICKNESS_FAULT[41] := BenchUut4.THICKNESS_FAULT;
   TraceIn_THICKNESS_SIGNAL_VALID[41] := BenchUut4.THICKNESS_SIGNAL_VALID;
   TraceIn_CUTTING_RUN[41] := BenchUut4.CUTTING_RUN;
   TraceIn_FaultTimestamp[41] := BenchUut4.FaultTimestamp;
   TraceIn_CycleTime[41] := BenchUut4.CycleTime;
   BenchUut4();
   TraceOut_THICKNESS_ALARM[41] := BenchUut4.THICKNESS_ALARM;
   TraceOut_Slab_Fault_Counter[41] := BenchUut4.Slab_Fault_Counter;
   TraceOut_Slab_Runtime_Accumulator[41] := BenchUut4.Slab_Runtime_Accumulator;
   TraceOut_Slab_Fault_History_0[41] := BenchUut4.Slab_Fault_History[0];
   TraceOut_Slab_Fault_History_1[41] := BenchUut4.Slab_Fault_History[1];
   TraceOut_Slab_Fault_History_2[41] := BenchUut4.Slab_Fault_History[2];
   TraceOut_Slab_Fault_History_3[41] := BenchUut4.Slab_Fault_History[3];
   TraceOut_Slab_Fault_History_4[41] := BenchUut4.Slab_Fault_History[4];
   BenchCalls := BenchCalls + 1;
   BenchStep := BenchStep + 1;
  END_IF;
 42:
  IF BenchCurrentTime - BenchLastTime >= UDINT_TO_TIME(300) THEN
   TraceDt[42] := TIME_TO_UDINT(BenchCurrentTime - BenchLastTime);
   BenchLastTime := BenchCurrentTime;
   BenchUut4.THICKNESS_FAULT := FALSE;
   BenchUut4.THICKNESS_SIGNAL_VALID := TRUE;
   BenchUut4.CUTTING_RUN := FALSE;
   BenchUut4.FaultTimestamp := DINT#20;
   BenchUut4.CycleTime := T#100ms;
   TraceIn_THICKNESS_FAULT[42] := BenchUut4.THICKNESS_FAULT;
   TraceIn_THICKNESS_SIGNAL_VALID[42] := BenchUut4.THICKNESS_SIGNAL_VALID;
   TraceIn_CUTTING_RUN[42] := BenchUut4.CUTTING_RUN;
   TraceIn_FaultTimestamp[42] := BenchUut4.FaultTimestamp;
   TraceIn_CycleTime[42] := BenchUut4.CycleTime;
   BenchUut4();
   TraceOut_THICKNESS_ALARM[42] := BenchUut4.THICKNESS_ALARM;
   TraceOut_Slab_Fault_Counter[42] := BenchUut4.Slab_Fault_Counter;
   TraceOut_Slab_Runtime_Accumulator[42] := BenchUut4.Slab_Runtime_Accumulator;
   TraceOut_Slab_Fault_History_0[42] := BenchUut4.Slab_Fault_History[0];
   TraceOut_Slab_Fault_History_1[42] := BenchUut4.Slab_Fault_History[1];
   TraceOut_Slab_Fault_History_2[42] := BenchUut4.Slab_Fault_History[2];
   TraceOut_Slab_Fault_History_3[42] := BenchUut4.Slab_Fault_History[3];
   TraceOut_Slab_Fault_History_4[42] := BenchUut4.Slab_Fault_History[4];
   BenchCalls := BenchCalls + 1;
   BenchStep := BenchStep + 1;
  END_IF;
 43:
  IF BenchCurrentTime - BenchLastTime >= UDINT_TO_TIME(200) THEN
   TraceDt[43] := TIME_TO_UDINT(BenchCurrentTime - BenchLastTime);
   BenchLastTime := BenchCurrentTime;
   BenchUut4.THICKNESS_FAULT := FALSE;
   BenchUut4.THICKNESS_SIGNAL_VALID := TRUE;
   BenchUut4.CUTTING_RUN := FALSE;
   BenchUut4.FaultTimestamp := DINT#20;
   BenchUut4.CycleTime := T#100ms;
   TraceIn_THICKNESS_FAULT[43] := BenchUut4.THICKNESS_FAULT;
   TraceIn_THICKNESS_SIGNAL_VALID[43] := BenchUut4.THICKNESS_SIGNAL_VALID;
   TraceIn_CUTTING_RUN[43] := BenchUut4.CUTTING_RUN;
   TraceIn_FaultTimestamp[43] := BenchUut4.FaultTimestamp;
   TraceIn_CycleTime[43] := BenchUut4.CycleTime;
   BenchUut4();
   TraceOut_THICKNESS_ALARM[43] := BenchUut4.THICKNESS_ALARM;
   TraceOut_Slab_Fault_Counter[43] := BenchUut4.Slab_Fault_Counter;
   TraceOut_Slab_Runtime_Accumulator[43] := BenchUut4.Slab_Runtime_Accumulator;
   TraceOut_Slab_Fault_History_0[43] := BenchUut4.Slab_Fault_History[0];
   TraceOut_Slab_Fault_History_1[43] := BenchUut4.Slab_Fault_History[1];
   TraceOut_Slab_Fault_History_2[43] := BenchUut4.Slab_Fault_History[2];
   TraceOut_Slab_Fault_History_3[43] := BenchUut4.Slab_Fault_History[3];
   TraceOut_Slab_Fault_History_4[43] := BenchUut4.Slab_Fault_History[4];
   BenchCalls := BenchCalls + 1;
   BenchStep := BenchStep + 1;
  END_IF;
 44:
  IF BenchCurrentTime - BenchLastTime >= UDINT_TO_TIME(100) THEN
   TraceDt[44] := TIME_TO_UDINT(BenchCurrentTime - BenchLastTime);
   BenchLastTime := BenchCurrentTime;
   BenchUut4.THICKNESS_FAULT := TRUE;
   BenchUut4.THICKNESS_SIGNAL_VALID := FALSE;
   BenchUut4.CUTTING_RUN := FALSE;
   BenchUut4.FaultTimestamp := DINT#20;
   BenchUut4.CycleTime := T#100ms;
   TraceIn_THICKNESS_FAULT[44] := BenchUut4.THICKNESS_FAULT;
   TraceIn_THICKNESS_SIGNAL_VALID[44] := BenchUut4.THICKNESS_SIGNAL_VALID;
   TraceIn_CUTTING_RUN[44] := BenchUut4.CUTTING_RUN;
   TraceIn_FaultTimestamp[44] := BenchUut4.FaultTimestamp;
   TraceIn_CycleTime[44] := BenchUut4.CycleTime;
   BenchUut4();
   TraceOut_THICKNESS_ALARM[44] := BenchUut4.THICKNESS_ALARM;
   TraceOut_Slab_Fault_Counter[44] := BenchUut4.Slab_Fault_Counter;
   TraceOut_Slab_Runtime_Accumulator[44] := BenchUut4.Slab_Runtime_Accumulator;
   TraceOut_Slab_Fault_History_0[44] := BenchUut4.Slab_Fault_History[0];
   TraceOut_Slab_Fault_History_1[44] := BenchUut4.Slab_Fault_History[1];
   TraceOut_Slab_Fault_History_2[44] := BenchUut4.Slab_Fault_History[2];
   TraceOut_Slab_Fault_History_3[44] := BenchUut4.Slab_Fault_History[3];
   TraceOut_Slab_Fault_History_4[44] := BenchUut4.Slab_Fault_History[4];
   BenchCalls := BenchCalls + 1;
   BenchStep := BenchStep + 1;
  END_IF;
 45:
  IF BenchCurrentTime - BenchLastTime >= UDINT_TO_TIME(100) THEN
   TraceDt[45] := TIME_TO_UDINT(BenchCurrentTime - BenchLastTime);
   BenchLastTime := BenchCurrentTime;
   BenchUut4.THICKNESS_FAULT := TRUE;
   BenchUut4.THICKNESS_SIGNAL_VALID := TRUE;
   BenchUut4.CUTTING_RUN := FALSE;
   BenchUut4.FaultTimestamp := DINT#30;
   BenchUut4.CycleTime := T#100ms;
   TraceIn_THICKNESS_FAULT[45] := BenchUut4.THICKNESS_FAULT;
   TraceIn_THICKNESS_SIGNAL_VALID[45] := BenchUut4.THICKNESS_SIGNAL_VALID;
   TraceIn_CUTTING_RUN[45] := BenchUut4.CUTTING_RUN;
   TraceIn_FaultTimestamp[45] := BenchUut4.FaultTimestamp;
   TraceIn_CycleTime[45] := BenchUut4.CycleTime;
   BenchUut4();
   TraceOut_THICKNESS_ALARM[45] := BenchUut4.THICKNESS_ALARM;
   TraceOut_Slab_Fault_Counter[45] := BenchUut4.Slab_Fault_Counter;
   TraceOut_Slab_Runtime_Accumulator[45] := BenchUut4.Slab_Runtime_Accumulator;
   TraceOut_Slab_Fault_History_0[45] := BenchUut4.Slab_Fault_History[0];
   TraceOut_Slab_Fault_History_1[45] := BenchUut4.Slab_Fault_History[1];
   TraceOut_Slab_Fault_History_2[45] := BenchUut4.Slab_Fault_History[2];
   TraceOut_Slab_Fault_History_3[45] := BenchUut4.Slab_Fault_History[3];
   TraceOut_Slab_Fault_History_4[45] := BenchUut4.Slab_Fault_History[4];
   BenchCalls := BenchCalls + 1;
   BenchStep := BenchStep + 1;
  END_IF;
 46:
  IF BenchCurrentTime - BenchLastTime >= UDINT_TO_TIME(100) THEN
   TraceDt[46] := TIME_TO_UDINT(BenchCurrentTime - BenchLastTime);
   BenchLastTime := BenchCurrentTime;
   BenchUut4.THICKNESS_FAULT := TRUE;
   BenchUut4.THICKNESS_SIGNAL_VALID := TRUE;
   BenchUut4.CUTTING_RUN := FALSE;
   BenchUut4.FaultTimestamp := DINT#30;
   BenchUut4.CycleTime := T#100ms;
   TraceIn_THICKNESS_FAULT[46] := BenchUut4.THICKNESS_FAULT;
   TraceIn_THICKNESS_SIGNAL_VALID[46] := BenchUut4.THICKNESS_SIGNAL_VALID;
   TraceIn_CUTTING_RUN[46] := BenchUut4.CUTTING_RUN;
   TraceIn_FaultTimestamp[46] := BenchUut4.FaultTimestamp;
   TraceIn_CycleTime[46] := BenchUut4.CycleTime;
   BenchUut4();
   TraceOut_THICKNESS_ALARM[46] := BenchUut4.THICKNESS_ALARM;
   TraceOut_Slab_Fault_Counter[46] := BenchUut4.Slab_Fault_Counter;
   TraceOut_Slab_Runtime_Accumulator[46] := BenchUut4.Slab_Runtime_Accumulator;
   TraceOut_Slab_Fault_History_0[46] := BenchUut4.Slab_Fault_History[0];
   TraceOut_Slab_Fault_History_1[46] := BenchUut4.Slab_Fault_History[1];
   TraceOut_Slab_Fault_History_2[46] := BenchUut4.Slab_Fault_History[2];
   TraceOut_Slab_Fault_History_3[46] := BenchUut4.Slab_Fault_History[3];
   TraceOut_Slab_Fault_History_4[46] := BenchUut4.Slab_Fault_History[4];
   BenchCalls := BenchCalls + 1;
   BenchStep := BenchStep + 1;
  END_IF;
 47:
  IF BenchCurrentTime - BenchLastTime >= UDINT_TO_TIME(0) THEN
   TraceDt[47] := TIME_TO_UDINT(BenchCurrentTime - BenchLastTime);
   BenchLastTime := BenchCurrentTime;
   BenchUut5.THICKNESS_FAULT := FALSE;
   BenchUut5.THICKNESS_SIGNAL_VALID := TRUE;
   BenchUut5.CUTTING_RUN := FALSE;
   BenchUut5.FaultTimestamp := DINT#0;
   BenchUut5.CycleTime := T#100ms;
   TraceIn_THICKNESS_FAULT[47] := BenchUut5.THICKNESS_FAULT;
   TraceIn_THICKNESS_SIGNAL_VALID[47] := BenchUut5.THICKNESS_SIGNAL_VALID;
   TraceIn_CUTTING_RUN[47] := BenchUut5.CUTTING_RUN;
   TraceIn_FaultTimestamp[47] := BenchUut5.FaultTimestamp;
   TraceIn_CycleTime[47] := BenchUut5.CycleTime;
   BenchUut5();
   TraceOut_THICKNESS_ALARM[47] := BenchUut5.THICKNESS_ALARM;
   TraceOut_Slab_Fault_Counter[47] := BenchUut5.Slab_Fault_Counter;
   TraceOut_Slab_Runtime_Accumulator[47] := BenchUut5.Slab_Runtime_Accumulator;
   TraceOut_Slab_Fault_History_0[47] := BenchUut5.Slab_Fault_History[0];
   TraceOut_Slab_Fault_History_1[47] := BenchUut5.Slab_Fault_History[1];
   TraceOut_Slab_Fault_History_2[47] := BenchUut5.Slab_Fault_History[2];
   TraceOut_Slab_Fault_History_3[47] := BenchUut5.Slab_Fault_History[3];
   TraceOut_Slab_Fault_History_4[47] := BenchUut5.Slab_Fault_History[4];
   BenchCalls := BenchCalls + 1;
   BenchStep := BenchStep + 1;
  END_IF;
 48:
  IF BenchCurrentTime - BenchLastTime >= UDINT_TO_TIME(100) THEN
   TraceDt[48] := TIME_TO_UDINT(BenchCurrentTime - BenchLastTime);
   BenchLastTime := BenchCurrentTime;
   BenchUut5.THICKNESS_FAULT := TRUE;
   BenchUut5.THICKNESS_SIGNAL_VALID := TRUE;
   BenchUut5.CUTTING_RUN := FALSE;
   BenchUut5.FaultTimestamp := DINT#101;
   BenchUut5.CycleTime := T#100ms;
   TraceIn_THICKNESS_FAULT[48] := BenchUut5.THICKNESS_FAULT;
   TraceIn_THICKNESS_SIGNAL_VALID[48] := BenchUut5.THICKNESS_SIGNAL_VALID;
   TraceIn_CUTTING_RUN[48] := BenchUut5.CUTTING_RUN;
   TraceIn_FaultTimestamp[48] := BenchUut5.FaultTimestamp;
   TraceIn_CycleTime[48] := BenchUut5.CycleTime;
   BenchUut5();
   TraceOut_THICKNESS_ALARM[48] := BenchUut5.THICKNESS_ALARM;
   TraceOut_Slab_Fault_Counter[48] := BenchUut5.Slab_Fault_Counter;
   TraceOut_Slab_Runtime_Accumulator[48] := BenchUut5.Slab_Runtime_Accumulator;
   TraceOut_Slab_Fault_History_0[48] := BenchUut5.Slab_Fault_History[0];
   TraceOut_Slab_Fault_History_1[48] := BenchUut5.Slab_Fault_History[1];
   TraceOut_Slab_Fault_History_2[48] := BenchUut5.Slab_Fault_History[2];
   TraceOut_Slab_Fault_History_3[48] := BenchUut5.Slab_Fault_History[3];
   TraceOut_Slab_Fault_History_4[48] := BenchUut5.Slab_Fault_History[4];
   BenchCalls := BenchCalls + 1;
   BenchStep := BenchStep + 1;
  END_IF;
 49:
  IF BenchCurrentTime - BenchLastTime >= UDINT_TO_TIME(100) THEN
   TraceDt[49] := TIME_TO_UDINT(BenchCurrentTime - BenchLastTime);
   BenchLastTime := BenchCurrentTime;
   BenchUut5.THICKNESS_FAULT := FALSE;
   BenchUut5.THICKNESS_SIGNAL_VALID := TRUE;
   BenchUut5.CUTTING_RUN := FALSE;
   BenchUut5.FaultTimestamp := DINT#0;
   BenchUut5.CycleTime := T#100ms;
   TraceIn_THICKNESS_FAULT[49] := BenchUut5.THICKNESS_FAULT;
   TraceIn_THICKNESS_SIGNAL_VALID[49] := BenchUut5.THICKNESS_SIGNAL_VALID;
   TraceIn_CUTTING_RUN[49] := BenchUut5.CUTTING_RUN;
   TraceIn_FaultTimestamp[49] := BenchUut5.FaultTimestamp;
   TraceIn_CycleTime[49] := BenchUut5.CycleTime;
   BenchUut5();
   TraceOut_THICKNESS_ALARM[49] := BenchUut5.THICKNESS_ALARM;
   TraceOut_Slab_Fault_Counter[49] := BenchUut5.Slab_Fault_Counter;
   TraceOut_Slab_Runtime_Accumulator[49] := BenchUut5.Slab_Runtime_Accumulator;
   TraceOut_Slab_Fault_History_0[49] := BenchUut5.Slab_Fault_History[0];
   TraceOut_Slab_Fault_History_1[49] := BenchUut5.Slab_Fault_History[1];
   TraceOut_Slab_Fault_History_2[49] := BenchUut5.Slab_Fault_History[2];
   TraceOut_Slab_Fault_History_3[49] := BenchUut5.Slab_Fault_History[3];
   TraceOut_Slab_Fault_History_4[49] := BenchUut5.Slab_Fault_History[4];
   BenchCalls := BenchCalls + 1;
   BenchStep := BenchStep + 1;
  END_IF;
 50:
  IF BenchCurrentTime - BenchLastTime >= UDINT_TO_TIME(100) THEN
   TraceDt[50] := TIME_TO_UDINT(BenchCurrentTime - BenchLastTime);
   BenchLastTime := BenchCurrentTime;
   BenchUut5.THICKNESS_FAULT := TRUE;
   BenchUut5.THICKNESS_SIGNAL_VALID := TRUE;
   BenchUut5.CUTTING_RUN := FALSE;
   BenchUut5.FaultTimestamp := DINT#102;
   BenchUut5.CycleTime := T#100ms;
   TraceIn_THICKNESS_FAULT[50] := BenchUut5.THICKNESS_FAULT;
   TraceIn_THICKNESS_SIGNAL_VALID[50] := BenchUut5.THICKNESS_SIGNAL_VALID;
   TraceIn_CUTTING_RUN[50] := BenchUut5.CUTTING_RUN;
   TraceIn_FaultTimestamp[50] := BenchUut5.FaultTimestamp;
   TraceIn_CycleTime[50] := BenchUut5.CycleTime;
   BenchUut5();
   TraceOut_THICKNESS_ALARM[50] := BenchUut5.THICKNESS_ALARM;
   TraceOut_Slab_Fault_Counter[50] := BenchUut5.Slab_Fault_Counter;
   TraceOut_Slab_Runtime_Accumulator[50] := BenchUut5.Slab_Runtime_Accumulator;
   TraceOut_Slab_Fault_History_0[50] := BenchUut5.Slab_Fault_History[0];
   TraceOut_Slab_Fault_History_1[50] := BenchUut5.Slab_Fault_History[1];
   TraceOut_Slab_Fault_History_2[50] := BenchUut5.Slab_Fault_History[2];
   TraceOut_Slab_Fault_History_3[50] := BenchUut5.Slab_Fault_History[3];
   TraceOut_Slab_Fault_History_4[50] := BenchUut5.Slab_Fault_History[4];
   BenchCalls := BenchCalls + 1;
   BenchStep := BenchStep + 1;
  END_IF;
 51:
  IF BenchCurrentTime - BenchLastTime >= UDINT_TO_TIME(100) THEN
   TraceDt[51] := TIME_TO_UDINT(BenchCurrentTime - BenchLastTime);
   BenchLastTime := BenchCurrentTime;
   BenchUut5.THICKNESS_FAULT := FALSE;
   BenchUut5.THICKNESS_SIGNAL_VALID := TRUE;
   BenchUut5.CUTTING_RUN := FALSE;
   BenchUut5.FaultTimestamp := DINT#0;
   BenchUut5.CycleTime := T#100ms;
   TraceIn_THICKNESS_FAULT[51] := BenchUut5.THICKNESS_FAULT;
   TraceIn_THICKNESS_SIGNAL_VALID[51] := BenchUut5.THICKNESS_SIGNAL_VALID;
   TraceIn_CUTTING_RUN[51] := BenchUut5.CUTTING_RUN;
   TraceIn_FaultTimestamp[51] := BenchUut5.FaultTimestamp;
   TraceIn_CycleTime[51] := BenchUut5.CycleTime;
   BenchUut5();
   TraceOut_THICKNESS_ALARM[51] := BenchUut5.THICKNESS_ALARM;
   TraceOut_Slab_Fault_Counter[51] := BenchUut5.Slab_Fault_Counter;
   TraceOut_Slab_Runtime_Accumulator[51] := BenchUut5.Slab_Runtime_Accumulator;
   TraceOut_Slab_Fault_History_0[51] := BenchUut5.Slab_Fault_History[0];
   TraceOut_Slab_Fault_History_1[51] := BenchUut5.Slab_Fault_History[1];
   TraceOut_Slab_Fault_History_2[51] := BenchUut5.Slab_Fault_History[2];
   TraceOut_Slab_Fault_History_3[51] := BenchUut5.Slab_Fault_History[3];
   TraceOut_Slab_Fault_History_4[51] := BenchUut5.Slab_Fault_History[4];
   BenchCalls := BenchCalls + 1;
   BenchStep := BenchStep + 1;
  END_IF;
 52:
  IF BenchCurrentTime - BenchLastTime >= UDINT_TO_TIME(100) THEN
   TraceDt[52] := TIME_TO_UDINT(BenchCurrentTime - BenchLastTime);
   BenchLastTime := BenchCurrentTime;
   BenchUut5.THICKNESS_FAULT := TRUE;
   BenchUut5.THICKNESS_SIGNAL_VALID := TRUE;
   BenchUut5.CUTTING_RUN := FALSE;
   BenchUut5.FaultTimestamp := DINT#103;
   BenchUut5.CycleTime := T#100ms;
   TraceIn_THICKNESS_FAULT[52] := BenchUut5.THICKNESS_FAULT;
   TraceIn_THICKNESS_SIGNAL_VALID[52] := BenchUut5.THICKNESS_SIGNAL_VALID;
   TraceIn_CUTTING_RUN[52] := BenchUut5.CUTTING_RUN;
   TraceIn_FaultTimestamp[52] := BenchUut5.FaultTimestamp;
   TraceIn_CycleTime[52] := BenchUut5.CycleTime;
   BenchUut5();
   TraceOut_THICKNESS_ALARM[52] := BenchUut5.THICKNESS_ALARM;
   TraceOut_Slab_Fault_Counter[52] := BenchUut5.Slab_Fault_Counter;
   TraceOut_Slab_Runtime_Accumulator[52] := BenchUut5.Slab_Runtime_Accumulator;
   TraceOut_Slab_Fault_History_0[52] := BenchUut5.Slab_Fault_History[0];
   TraceOut_Slab_Fault_History_1[52] := BenchUut5.Slab_Fault_History[1];
   TraceOut_Slab_Fault_History_2[52] := BenchUut5.Slab_Fault_History[2];
   TraceOut_Slab_Fault_History_3[52] := BenchUut5.Slab_Fault_History[3];
   TraceOut_Slab_Fault_History_4[52] := BenchUut5.Slab_Fault_History[4];
   BenchCalls := BenchCalls + 1;
   BenchStep := BenchStep + 1;
  END_IF;
 53:
  IF BenchCurrentTime - BenchLastTime >= UDINT_TO_TIME(100) THEN
   TraceDt[53] := TIME_TO_UDINT(BenchCurrentTime - BenchLastTime);
   BenchLastTime := BenchCurrentTime;
   BenchUut5.THICKNESS_FAULT := FALSE;
   BenchUut5.THICKNESS_SIGNAL_VALID := TRUE;
   BenchUut5.CUTTING_RUN := FALSE;
   BenchUut5.FaultTimestamp := DINT#0;
   BenchUut5.CycleTime := T#100ms;
   TraceIn_THICKNESS_FAULT[53] := BenchUut5.THICKNESS_FAULT;
   TraceIn_THICKNESS_SIGNAL_VALID[53] := BenchUut5.THICKNESS_SIGNAL_VALID;
   TraceIn_CUTTING_RUN[53] := BenchUut5.CUTTING_RUN;
   TraceIn_FaultTimestamp[53] := BenchUut5.FaultTimestamp;
   TraceIn_CycleTime[53] := BenchUut5.CycleTime;
   BenchUut5();
   TraceOut_THICKNESS_ALARM[53] := BenchUut5.THICKNESS_ALARM;
   TraceOut_Slab_Fault_Counter[53] := BenchUut5.Slab_Fault_Counter;
   TraceOut_Slab_Runtime_Accumulator[53] := BenchUut5.Slab_Runtime_Accumulator;
   TraceOut_Slab_Fault_History_0[53] := BenchUut5.Slab_Fault_History[0];
   TraceOut_Slab_Fault_History_1[53] := BenchUut5.Slab_Fault_History[1];
   TraceOut_Slab_Fault_History_2[53] := BenchUut5.Slab_Fault_History[2];
   TraceOut_Slab_Fault_History_3[53] := BenchUut5.Slab_Fault_History[3];
   TraceOut_Slab_Fault_History_4[53] := BenchUut5.Slab_Fault_History[4];
   BenchCalls := BenchCalls + 1;
   BenchStep := BenchStep + 1;
  END_IF;
 54:
  IF BenchCurrentTime - BenchLastTime >= UDINT_TO_TIME(100) THEN
   TraceDt[54] := TIME_TO_UDINT(BenchCurrentTime - BenchLastTime);
   BenchLastTime := BenchCurrentTime;
   BenchUut5.THICKNESS_FAULT := TRUE;
   BenchUut5.THICKNESS_SIGNAL_VALID := TRUE;
   BenchUut5.CUTTING_RUN := FALSE;
   BenchUut5.FaultTimestamp := DINT#104;
   BenchUut5.CycleTime := T#100ms;
   TraceIn_THICKNESS_FAULT[54] := BenchUut5.THICKNESS_FAULT;
   TraceIn_THICKNESS_SIGNAL_VALID[54] := BenchUut5.THICKNESS_SIGNAL_VALID;
   TraceIn_CUTTING_RUN[54] := BenchUut5.CUTTING_RUN;
   TraceIn_FaultTimestamp[54] := BenchUut5.FaultTimestamp;
   TraceIn_CycleTime[54] := BenchUut5.CycleTime;
   BenchUut5();
   TraceOut_THICKNESS_ALARM[54] := BenchUut5.THICKNESS_ALARM;
   TraceOut_Slab_Fault_Counter[54] := BenchUut5.Slab_Fault_Counter;
   TraceOut_Slab_Runtime_Accumulator[54] := BenchUut5.Slab_Runtime_Accumulator;
   TraceOut_Slab_Fault_History_0[54] := BenchUut5.Slab_Fault_History[0];
   TraceOut_Slab_Fault_History_1[54] := BenchUut5.Slab_Fault_History[1];
   TraceOut_Slab_Fault_History_2[54] := BenchUut5.Slab_Fault_History[2];
   TraceOut_Slab_Fault_History_3[54] := BenchUut5.Slab_Fault_History[3];
   TraceOut_Slab_Fault_History_4[54] := BenchUut5.Slab_Fault_History[4];
   BenchCalls := BenchCalls + 1;
   BenchStep := BenchStep + 1;
  END_IF;
 55:
  IF BenchCurrentTime - BenchLastTime >= UDINT_TO_TIME(100) THEN
   TraceDt[55] := TIME_TO_UDINT(BenchCurrentTime - BenchLastTime);
   BenchLastTime := BenchCurrentTime;
   BenchUut5.THICKNESS_FAULT := FALSE;
   BenchUut5.THICKNESS_SIGNAL_VALID := TRUE;
   BenchUut5.CUTTING_RUN := FALSE;
   BenchUut5.FaultTimestamp := DINT#0;
   BenchUut5.CycleTime := T#100ms;
   TraceIn_THICKNESS_FAULT[55] := BenchUut5.THICKNESS_FAULT;
   TraceIn_THICKNESS_SIGNAL_VALID[55] := BenchUut5.THICKNESS_SIGNAL_VALID;
   TraceIn_CUTTING_RUN[55] := BenchUut5.CUTTING_RUN;
   TraceIn_FaultTimestamp[55] := BenchUut5.FaultTimestamp;
   TraceIn_CycleTime[55] := BenchUut5.CycleTime;
   BenchUut5();
   TraceOut_THICKNESS_ALARM[55] := BenchUut5.THICKNESS_ALARM;
   TraceOut_Slab_Fault_Counter[55] := BenchUut5.Slab_Fault_Counter;
   TraceOut_Slab_Runtime_Accumulator[55] := BenchUut5.Slab_Runtime_Accumulator;
   TraceOut_Slab_Fault_History_0[55] := BenchUut5.Slab_Fault_History[0];
   TraceOut_Slab_Fault_History_1[55] := BenchUut5.Slab_Fault_History[1];
   TraceOut_Slab_Fault_History_2[55] := BenchUut5.Slab_Fault_History[2];
   TraceOut_Slab_Fault_History_3[55] := BenchUut5.Slab_Fault_History[3];
   TraceOut_Slab_Fault_History_4[55] := BenchUut5.Slab_Fault_History[4];
   BenchCalls := BenchCalls + 1;
   BenchStep := BenchStep + 1;
  END_IF;
 56:
  IF BenchCurrentTime - BenchLastTime >= UDINT_TO_TIME(100) THEN
   TraceDt[56] := TIME_TO_UDINT(BenchCurrentTime - BenchLastTime);
   BenchLastTime := BenchCurrentTime;
   BenchUut5.THICKNESS_FAULT := TRUE;
   BenchUut5.THICKNESS_SIGNAL_VALID := TRUE;
   BenchUut5.CUTTING_RUN := FALSE;
   BenchUut5.FaultTimestamp := DINT#105;
   BenchUut5.CycleTime := T#100ms;
   TraceIn_THICKNESS_FAULT[56] := BenchUut5.THICKNESS_FAULT;
   TraceIn_THICKNESS_SIGNAL_VALID[56] := BenchUut5.THICKNESS_SIGNAL_VALID;
   TraceIn_CUTTING_RUN[56] := BenchUut5.CUTTING_RUN;
   TraceIn_FaultTimestamp[56] := BenchUut5.FaultTimestamp;
   TraceIn_CycleTime[56] := BenchUut5.CycleTime;
   BenchUut5();
   TraceOut_THICKNESS_ALARM[56] := BenchUut5.THICKNESS_ALARM;
   TraceOut_Slab_Fault_Counter[56] := BenchUut5.Slab_Fault_Counter;
   TraceOut_Slab_Runtime_Accumulator[56] := BenchUut5.Slab_Runtime_Accumulator;
   TraceOut_Slab_Fault_History_0[56] := BenchUut5.Slab_Fault_History[0];
   TraceOut_Slab_Fault_History_1[56] := BenchUut5.Slab_Fault_History[1];
   TraceOut_Slab_Fault_History_2[56] := BenchUut5.Slab_Fault_History[2];
   TraceOut_Slab_Fault_History_3[56] := BenchUut5.Slab_Fault_History[3];
   TraceOut_Slab_Fault_History_4[56] := BenchUut5.Slab_Fault_History[4];
   BenchCalls := BenchCalls + 1;
   BenchStep := BenchStep + 1;
  END_IF;
 57:
  IF BenchCurrentTime - BenchLastTime >= UDINT_TO_TIME(100) THEN
   TraceDt[57] := TIME_TO_UDINT(BenchCurrentTime - BenchLastTime);
   BenchLastTime := BenchCurrentTime;
   BenchUut5.THICKNESS_FAULT := FALSE;
   BenchUut5.THICKNESS_SIGNAL_VALID := TRUE;
   BenchUut5.CUTTING_RUN := FALSE;
   BenchUut5.FaultTimestamp := DINT#0;
   BenchUut5.CycleTime := T#100ms;
   TraceIn_THICKNESS_FAULT[57] := BenchUut5.THICKNESS_FAULT;
   TraceIn_THICKNESS_SIGNAL_VALID[57] := BenchUut5.THICKNESS_SIGNAL_VALID;
   TraceIn_CUTTING_RUN[57] := BenchUut5.CUTTING_RUN;
   TraceIn_FaultTimestamp[57] := BenchUut5.FaultTimestamp;
   TraceIn_CycleTime[57] := BenchUut5.CycleTime;
   BenchUut5();
   TraceOut_THICKNESS_ALARM[57] := BenchUut5.THICKNESS_ALARM;
   TraceOut_Slab_Fault_Counter[57] := BenchUut5.Slab_Fault_Counter;
   TraceOut_Slab_Runtime_Accumulator[57] := BenchUut5.Slab_Runtime_Accumulator;
   TraceOut_Slab_Fault_History_0[57] := BenchUut5.Slab_Fault_History[0];
   TraceOut_Slab_Fault_History_1[57] := BenchUut5.Slab_Fault_History[1];
   TraceOut_Slab_Fault_History_2[57] := BenchUut5.Slab_Fault_History[2];
   TraceOut_Slab_Fault_History_3[57] := BenchUut5.Slab_Fault_History[3];
   TraceOut_Slab_Fault_History_4[57] := BenchUut5.Slab_Fault_History[4];
   BenchCalls := BenchCalls + 1;
   BenchStep := BenchStep + 1;
  END_IF;
 58:
  IF BenchCurrentTime - BenchLastTime >= UDINT_TO_TIME(100) THEN
   TraceDt[58] := TIME_TO_UDINT(BenchCurrentTime - BenchLastTime);
   BenchLastTime := BenchCurrentTime;
   BenchUut5.THICKNESS_FAULT := TRUE;
   BenchUut5.THICKNESS_SIGNAL_VALID := TRUE;
   BenchUut5.CUTTING_RUN := FALSE;
   BenchUut5.FaultTimestamp := DINT#106;
   BenchUut5.CycleTime := T#100ms;
   TraceIn_THICKNESS_FAULT[58] := BenchUut5.THICKNESS_FAULT;
   TraceIn_THICKNESS_SIGNAL_VALID[58] := BenchUut5.THICKNESS_SIGNAL_VALID;
   TraceIn_CUTTING_RUN[58] := BenchUut5.CUTTING_RUN;
   TraceIn_FaultTimestamp[58] := BenchUut5.FaultTimestamp;
   TraceIn_CycleTime[58] := BenchUut5.CycleTime;
   BenchUut5();
   TraceOut_THICKNESS_ALARM[58] := BenchUut5.THICKNESS_ALARM;
   TraceOut_Slab_Fault_Counter[58] := BenchUut5.Slab_Fault_Counter;
   TraceOut_Slab_Runtime_Accumulator[58] := BenchUut5.Slab_Runtime_Accumulator;
   TraceOut_Slab_Fault_History_0[58] := BenchUut5.Slab_Fault_History[0];
   TraceOut_Slab_Fault_History_1[58] := BenchUut5.Slab_Fault_History[1];
   TraceOut_Slab_Fault_History_2[58] := BenchUut5.Slab_Fault_History[2];
   TraceOut_Slab_Fault_History_3[58] := BenchUut5.Slab_Fault_History[3];
   TraceOut_Slab_Fault_History_4[58] := BenchUut5.Slab_Fault_History[4];
   BenchCalls := BenchCalls + 1;
   BenchStep := BenchStep + 1;
  END_IF;
 59:
  IF BenchCurrentTime - BenchLastTime >= UDINT_TO_TIME(100) THEN
   TraceDt[59] := TIME_TO_UDINT(BenchCurrentTime - BenchLastTime);
   BenchLastTime := BenchCurrentTime;
   BenchUut5.THICKNESS_FAULT := FALSE;
   BenchUut5.THICKNESS_SIGNAL_VALID := TRUE;
   BenchUut5.CUTTING_RUN := FALSE;
   BenchUut5.FaultTimestamp := DINT#0;
   BenchUut5.CycleTime := T#100ms;
   TraceIn_THICKNESS_FAULT[59] := BenchUut5.THICKNESS_FAULT;
   TraceIn_THICKNESS_SIGNAL_VALID[59] := BenchUut5.THICKNESS_SIGNAL_VALID;
   TraceIn_CUTTING_RUN[59] := BenchUut5.CUTTING_RUN;
   TraceIn_FaultTimestamp[59] := BenchUut5.FaultTimestamp;
   TraceIn_CycleTime[59] := BenchUut5.CycleTime;
   BenchUut5();
   TraceOut_THICKNESS_ALARM[59] := BenchUut5.THICKNESS_ALARM;
   TraceOut_Slab_Fault_Counter[59] := BenchUut5.Slab_Fault_Counter;
   TraceOut_Slab_Runtime_Accumulator[59] := BenchUut5.Slab_Runtime_Accumulator;
   TraceOut_Slab_Fault_History_0[59] := BenchUut5.Slab_Fault_History[0];
   TraceOut_Slab_Fault_History_1[59] := BenchUut5.Slab_Fault_History[1];
   TraceOut_Slab_Fault_History_2[59] := BenchUut5.Slab_Fault_History[2];
   TraceOut_Slab_Fault_History_3[59] := BenchUut5.Slab_Fault_History[3];
   TraceOut_Slab_Fault_History_4[59] := BenchUut5.Slab_Fault_History[4];
   BenchCalls := BenchCalls + 1;
   BenchStep := BenchStep + 1;
  END_IF;
 60:
  IF BenchCurrentTime - BenchLastTime >= UDINT_TO_TIME(100) THEN
   TraceDt[60] := TIME_TO_UDINT(BenchCurrentTime - BenchLastTime);
   BenchLastTime := BenchCurrentTime;
   BenchUut5.THICKNESS_FAULT := TRUE;
   BenchUut5.THICKNESS_SIGNAL_VALID := TRUE;
   BenchUut5.CUTTING_RUN := FALSE;
   BenchUut5.FaultTimestamp := DINT#107;
   BenchUut5.CycleTime := T#100ms;
   TraceIn_THICKNESS_FAULT[60] := BenchUut5.THICKNESS_FAULT;
   TraceIn_THICKNESS_SIGNAL_VALID[60] := BenchUut5.THICKNESS_SIGNAL_VALID;
   TraceIn_CUTTING_RUN[60] := BenchUut5.CUTTING_RUN;
   TraceIn_FaultTimestamp[60] := BenchUut5.FaultTimestamp;
   TraceIn_CycleTime[60] := BenchUut5.CycleTime;
   BenchUut5();
   TraceOut_THICKNESS_ALARM[60] := BenchUut5.THICKNESS_ALARM;
   TraceOut_Slab_Fault_Counter[60] := BenchUut5.Slab_Fault_Counter;
   TraceOut_Slab_Runtime_Accumulator[60] := BenchUut5.Slab_Runtime_Accumulator;
   TraceOut_Slab_Fault_History_0[60] := BenchUut5.Slab_Fault_History[0];
   TraceOut_Slab_Fault_History_1[60] := BenchUut5.Slab_Fault_History[1];
   TraceOut_Slab_Fault_History_2[60] := BenchUut5.Slab_Fault_History[2];
   TraceOut_Slab_Fault_History_3[60] := BenchUut5.Slab_Fault_History[3];
   TraceOut_Slab_Fault_History_4[60] := BenchUut5.Slab_Fault_History[4];
   BenchCalls := BenchCalls + 1;
   BenchStep := BenchStep + 1;
  END_IF;
 61:
  IF BenchCurrentTime - BenchLastTime >= UDINT_TO_TIME(0) THEN
   TraceDt[61] := TIME_TO_UDINT(BenchCurrentTime - BenchLastTime);
   BenchLastTime := BenchCurrentTime;
   BenchUut6.THICKNESS_FAULT := FALSE;
   BenchUut6.THICKNESS_SIGNAL_VALID := TRUE;
   BenchUut6.CUTTING_RUN := TRUE;
   BenchUut6.FaultTimestamp := DINT#0;
   BenchUut6.CycleTime := T#200ms;
   TraceIn_THICKNESS_FAULT[61] := BenchUut6.THICKNESS_FAULT;
   TraceIn_THICKNESS_SIGNAL_VALID[61] := BenchUut6.THICKNESS_SIGNAL_VALID;
   TraceIn_CUTTING_RUN[61] := BenchUut6.CUTTING_RUN;
   TraceIn_FaultTimestamp[61] := BenchUut6.FaultTimestamp;
   TraceIn_CycleTime[61] := BenchUut6.CycleTime;
   BenchUut6();
   TraceOut_THICKNESS_ALARM[61] := BenchUut6.THICKNESS_ALARM;
   TraceOut_Slab_Fault_Counter[61] := BenchUut6.Slab_Fault_Counter;
   TraceOut_Slab_Runtime_Accumulator[61] := BenchUut6.Slab_Runtime_Accumulator;
   TraceOut_Slab_Fault_History_0[61] := BenchUut6.Slab_Fault_History[0];
   TraceOut_Slab_Fault_History_1[61] := BenchUut6.Slab_Fault_History[1];
   TraceOut_Slab_Fault_History_2[61] := BenchUut6.Slab_Fault_History[2];
   TraceOut_Slab_Fault_History_3[61] := BenchUut6.Slab_Fault_History[3];
   TraceOut_Slab_Fault_History_4[61] := BenchUut6.Slab_Fault_History[4];
   BenchCalls := BenchCalls + 1;
   BenchStep := BenchStep + 1;
  END_IF;
 62:
  IF BenchCurrentTime - BenchLastTime >= UDINT_TO_TIME(200) THEN
   TraceDt[62] := TIME_TO_UDINT(BenchCurrentTime - BenchLastTime);
   BenchLastTime := BenchCurrentTime;
   BenchUut6.THICKNESS_FAULT := TRUE;
   BenchUut6.THICKNESS_SIGNAL_VALID := FALSE;
   BenchUut6.CUTTING_RUN := TRUE;
   BenchUut6.FaultTimestamp := DINT#555;
   BenchUut6.CycleTime := T#200ms;
   TraceIn_THICKNESS_FAULT[62] := BenchUut6.THICKNESS_FAULT;
   TraceIn_THICKNESS_SIGNAL_VALID[62] := BenchUut6.THICKNESS_SIGNAL_VALID;
   TraceIn_CUTTING_RUN[62] := BenchUut6.CUTTING_RUN;
   TraceIn_FaultTimestamp[62] := BenchUut6.FaultTimestamp;
   TraceIn_CycleTime[62] := BenchUut6.CycleTime;
   BenchUut6();
   TraceOut_THICKNESS_ALARM[62] := BenchUut6.THICKNESS_ALARM;
   TraceOut_Slab_Fault_Counter[62] := BenchUut6.Slab_Fault_Counter;
   TraceOut_Slab_Runtime_Accumulator[62] := BenchUut6.Slab_Runtime_Accumulator;
   TraceOut_Slab_Fault_History_0[62] := BenchUut6.Slab_Fault_History[0];
   TraceOut_Slab_Fault_History_1[62] := BenchUut6.Slab_Fault_History[1];
   TraceOut_Slab_Fault_History_2[62] := BenchUut6.Slab_Fault_History[2];
   TraceOut_Slab_Fault_History_3[62] := BenchUut6.Slab_Fault_History[3];
   TraceOut_Slab_Fault_History_4[62] := BenchUut6.Slab_Fault_History[4];
   BenchCalls := BenchCalls + 1;
   BenchStep := BenchStep + 1;
  END_IF;
 63:
  IF BenchCurrentTime - BenchLastTime >= UDINT_TO_TIME(200) THEN
   TraceDt[63] := TIME_TO_UDINT(BenchCurrentTime - BenchLastTime);
   BenchLastTime := BenchCurrentTime;
   BenchUut6.THICKNESS_FAULT := TRUE;
   BenchUut6.THICKNESS_SIGNAL_VALID := TRUE;
   BenchUut6.CUTTING_RUN := TRUE;
   BenchUut6.FaultTimestamp := DINT#777;
   BenchUut6.CycleTime := T#200ms;
   TraceIn_THICKNESS_FAULT[63] := BenchUut6.THICKNESS_FAULT;
   TraceIn_THICKNESS_SIGNAL_VALID[63] := BenchUut6.THICKNESS_SIGNAL_VALID;
   TraceIn_CUTTING_RUN[63] := BenchUut6.CUTTING_RUN;
   TraceIn_FaultTimestamp[63] := BenchUut6.FaultTimestamp;
   TraceIn_CycleTime[63] := BenchUut6.CycleTime;
   BenchUut6();
   TraceOut_THICKNESS_ALARM[63] := BenchUut6.THICKNESS_ALARM;
   TraceOut_Slab_Fault_Counter[63] := BenchUut6.Slab_Fault_Counter;
   TraceOut_Slab_Runtime_Accumulator[63] := BenchUut6.Slab_Runtime_Accumulator;
   TraceOut_Slab_Fault_History_0[63] := BenchUut6.Slab_Fault_History[0];
   TraceOut_Slab_Fault_History_1[63] := BenchUut6.Slab_Fault_History[1];
   TraceOut_Slab_Fault_History_2[63] := BenchUut6.Slab_Fault_History[2];
   TraceOut_Slab_Fault_History_3[63] := BenchUut6.Slab_Fault_History[3];
   TraceOut_Slab_Fault_History_4[63] := BenchUut6.Slab_Fault_History[4];
   BenchCalls := BenchCalls + 1;
   BenchStep := BenchStep + 1;
  END_IF;
 64:
  IF BenchCurrentTime - BenchLastTime >= UDINT_TO_TIME(200) THEN
   TraceDt[64] := TIME_TO_UDINT(BenchCurrentTime - BenchLastTime);
   BenchLastTime := BenchCurrentTime;
   BenchUut6.THICKNESS_FAULT := FALSE;
   BenchUut6.THICKNESS_SIGNAL_VALID := TRUE;
   BenchUut6.CUTTING_RUN := TRUE;
   BenchUut6.FaultTimestamp := DINT#0;
   BenchUut6.CycleTime := T#200ms;
   TraceIn_THICKNESS_FAULT[64] := BenchUut6.THICKNESS_FAULT;
   TraceIn_THICKNESS_SIGNAL_VALID[64] := BenchUut6.THICKNESS_SIGNAL_VALID;
   TraceIn_CUTTING_RUN[64] := BenchUut6.CUTTING_RUN;
   TraceIn_FaultTimestamp[64] := BenchUut6.FaultTimestamp;
   TraceIn_CycleTime[64] := BenchUut6.CycleTime;
   BenchUut6();
   TraceOut_THICKNESS_ALARM[64] := BenchUut6.THICKNESS_ALARM;
   TraceOut_Slab_Fault_Counter[64] := BenchUut6.Slab_Fault_Counter;
   TraceOut_Slab_Runtime_Accumulator[64] := BenchUut6.Slab_Runtime_Accumulator;
   TraceOut_Slab_Fault_History_0[64] := BenchUut6.Slab_Fault_History[0];
   TraceOut_Slab_Fault_History_1[64] := BenchUut6.Slab_Fault_History[1];
   TraceOut_Slab_Fault_History_2[64] := BenchUut6.Slab_Fault_History[2];
   TraceOut_Slab_Fault_History_3[64] := BenchUut6.Slab_Fault_History[3];
   TraceOut_Slab_Fault_History_4[64] := BenchUut6.Slab_Fault_History[4];
   BenchCalls := BenchCalls + 1;
   BenchStep := BenchStep + 1;
  END_IF;
 65:
  IF BenchCurrentTime - BenchLastTime >= UDINT_TO_TIME(200) THEN
   TraceDt[65] := TIME_TO_UDINT(BenchCurrentTime - BenchLastTime);
   BenchLastTime := BenchCurrentTime;
   BenchUut6.THICKNESS_FAULT := FALSE;
   BenchUut6.THICKNESS_SIGNAL_VALID := TRUE;
   BenchUut6.CUTTING_RUN := FALSE;
   BenchUut6.FaultTimestamp := DINT#0;
   BenchUut6.CycleTime := T#200ms;
   TraceIn_THICKNESS_FAULT[65] := BenchUut6.THICKNESS_FAULT;
   TraceIn_THICKNESS_SIGNAL_VALID[65] := BenchUut6.THICKNESS_SIGNAL_VALID;
   TraceIn_CUTTING_RUN[65] := BenchUut6.CUTTING_RUN;
   TraceIn_FaultTimestamp[65] := BenchUut6.FaultTimestamp;
   TraceIn_CycleTime[65] := BenchUut6.CycleTime;
   BenchUut6();
   TraceOut_THICKNESS_ALARM[65] := BenchUut6.THICKNESS_ALARM;
   TraceOut_Slab_Fault_Counter[65] := BenchUut6.Slab_Fault_Counter;
   TraceOut_Slab_Runtime_Accumulator[65] := BenchUut6.Slab_Runtime_Accumulator;
   TraceOut_Slab_Fault_History_0[65] := BenchUut6.Slab_Fault_History[0];
   TraceOut_Slab_Fault_History_1[65] := BenchUut6.Slab_Fault_History[1];
   TraceOut_Slab_Fault_History_2[65] := BenchUut6.Slab_Fault_History[2];
   TraceOut_Slab_Fault_History_3[65] := BenchUut6.Slab_Fault_History[3];
   TraceOut_Slab_Fault_History_4[65] := BenchUut6.Slab_Fault_History[4];
   BenchCalls := BenchCalls + 1;
   BenchStep := BenchStep + 1;
  END_IF;
 66:
  IF BenchCurrentTime - BenchLastTime >= UDINT_TO_TIME(0) THEN
   TraceDt[66] := TIME_TO_UDINT(BenchCurrentTime - BenchLastTime);
   BenchLastTime := BenchCurrentTime;
   BenchUut7.THICKNESS_FAULT := TRUE;
   BenchUut7.THICKNESS_SIGNAL_VALID := TRUE;
   BenchUut7.CUTTING_RUN := FALSE;
   BenchUut7.FaultTimestamp := DINT#900;
   BenchUut7.CycleTime := T#100ms;
   TraceIn_THICKNESS_FAULT[66] := BenchUut7.THICKNESS_FAULT;
   TraceIn_THICKNESS_SIGNAL_VALID[66] := BenchUut7.THICKNESS_SIGNAL_VALID;
   TraceIn_CUTTING_RUN[66] := BenchUut7.CUTTING_RUN;
   TraceIn_FaultTimestamp[66] := BenchUut7.FaultTimestamp;
   TraceIn_CycleTime[66] := BenchUut7.CycleTime;
   BenchUut7();
   TraceOut_THICKNESS_ALARM[66] := BenchUut7.THICKNESS_ALARM;
   TraceOut_Slab_Fault_Counter[66] := BenchUut7.Slab_Fault_Counter;
   TraceOut_Slab_Runtime_Accumulator[66] := BenchUut7.Slab_Runtime_Accumulator;
   TraceOut_Slab_Fault_History_0[66] := BenchUut7.Slab_Fault_History[0];
   TraceOut_Slab_Fault_History_1[66] := BenchUut7.Slab_Fault_History[1];
   TraceOut_Slab_Fault_History_2[66] := BenchUut7.Slab_Fault_History[2];
   TraceOut_Slab_Fault_History_3[66] := BenchUut7.Slab_Fault_History[3];
   TraceOut_Slab_Fault_History_4[66] := BenchUut7.Slab_Fault_History[4];
   BenchCalls := BenchCalls + 1;
   BenchStep := BenchStep + 1;
  END_IF;
 67:
  IF BenchCurrentTime - BenchLastTime >= UDINT_TO_TIME(100) THEN
   TraceDt[67] := TIME_TO_UDINT(BenchCurrentTime - BenchLastTime);
   BenchLastTime := BenchCurrentTime;
   BenchUut7.THICKNESS_FAULT := TRUE;
   BenchUut7.THICKNESS_SIGNAL_VALID := TRUE;
   BenchUut7.CUTTING_RUN := FALSE;
   BenchUut7.FaultTimestamp := DINT#901;
   BenchUut7.CycleTime := T#100ms;
   TraceIn_THICKNESS_FAULT[67] := BenchUut7.THICKNESS_FAULT;
   TraceIn_THICKNESS_SIGNAL_VALID[67] := BenchUut7.THICKNESS_SIGNAL_VALID;
   TraceIn_CUTTING_RUN[67] := BenchUut7.CUTTING_RUN;
   TraceIn_FaultTimestamp[67] := BenchUut7.FaultTimestamp;
   TraceIn_CycleTime[67] := BenchUut7.CycleTime;
   BenchUut7();
   TraceOut_THICKNESS_ALARM[67] := BenchUut7.THICKNESS_ALARM;
   TraceOut_Slab_Fault_Counter[67] := BenchUut7.Slab_Fault_Counter;
   TraceOut_Slab_Runtime_Accumulator[67] := BenchUut7.Slab_Runtime_Accumulator;
   TraceOut_Slab_Fault_History_0[67] := BenchUut7.Slab_Fault_History[0];
   TraceOut_Slab_Fault_History_1[67] := BenchUut7.Slab_Fault_History[1];
   TraceOut_Slab_Fault_History_2[67] := BenchUut7.Slab_Fault_History[2];
   TraceOut_Slab_Fault_History_3[67] := BenchUut7.Slab_Fault_History[3];
   TraceOut_Slab_Fault_History_4[67] := BenchUut7.Slab_Fault_History[4];
   BenchCalls := BenchCalls + 1;
   BenchStep := BenchStep + 1;
  END_IF;
 68:
  IF BenchCurrentTime - BenchLastTime >= UDINT_TO_TIME(399) THEN
   TraceDt[68] := TIME_TO_UDINT(BenchCurrentTime - BenchLastTime);
   BenchLastTime := BenchCurrentTime;
   BenchUut7.THICKNESS_FAULT := FALSE;
   BenchUut7.THICKNESS_SIGNAL_VALID := TRUE;
   BenchUut7.CUTTING_RUN := FALSE;
   BenchUut7.FaultTimestamp := DINT#0;
   BenchUut7.CycleTime := T#100ms;
   TraceIn_THICKNESS_FAULT[68] := BenchUut7.THICKNESS_FAULT;
   TraceIn_THICKNESS_SIGNAL_VALID[68] := BenchUut7.THICKNESS_SIGNAL_VALID;
   TraceIn_CUTTING_RUN[68] := BenchUut7.CUTTING_RUN;
   TraceIn_FaultTimestamp[68] := BenchUut7.FaultTimestamp;
   TraceIn_CycleTime[68] := BenchUut7.CycleTime;
   BenchUut7();
   TraceOut_THICKNESS_ALARM[68] := BenchUut7.THICKNESS_ALARM;
   TraceOut_Slab_Fault_Counter[68] := BenchUut7.Slab_Fault_Counter;
   TraceOut_Slab_Runtime_Accumulator[68] := BenchUut7.Slab_Runtime_Accumulator;
   TraceOut_Slab_Fault_History_0[68] := BenchUut7.Slab_Fault_History[0];
   TraceOut_Slab_Fault_History_1[68] := BenchUut7.Slab_Fault_History[1];
   TraceOut_Slab_Fault_History_2[68] := BenchUut7.Slab_Fault_History[2];
   TraceOut_Slab_Fault_History_3[68] := BenchUut7.Slab_Fault_History[3];
   TraceOut_Slab_Fault_History_4[68] := BenchUut7.Slab_Fault_History[4];
   BenchCalls := BenchCalls + 1;
   BenchStep := BenchStep + 1;
  END_IF;
 69:
  IF BenchCurrentTime - BenchLastTime >= UDINT_TO_TIME(1) THEN
   TraceDt[69] := TIME_TO_UDINT(BenchCurrentTime - BenchLastTime);
   BenchLastTime := BenchCurrentTime;
   BenchUut7.THICKNESS_FAULT := FALSE;
   BenchUut7.THICKNESS_SIGNAL_VALID := TRUE;
   BenchUut7.CUTTING_RUN := FALSE;
   BenchUut7.FaultTimestamp := DINT#0;
   BenchUut7.CycleTime := T#100ms;
   TraceIn_THICKNESS_FAULT[69] := BenchUut7.THICKNESS_FAULT;
   TraceIn_THICKNESS_SIGNAL_VALID[69] := BenchUut7.THICKNESS_SIGNAL_VALID;
   TraceIn_CUTTING_RUN[69] := BenchUut7.CUTTING_RUN;
   TraceIn_FaultTimestamp[69] := BenchUut7.FaultTimestamp;
   TraceIn_CycleTime[69] := BenchUut7.CycleTime;
   BenchUut7();
   TraceOut_THICKNESS_ALARM[69] := BenchUut7.THICKNESS_ALARM;
   TraceOut_Slab_Fault_Counter[69] := BenchUut7.Slab_Fault_Counter;
   TraceOut_Slab_Runtime_Accumulator[69] := BenchUut7.Slab_Runtime_Accumulator;
   TraceOut_Slab_Fault_History_0[69] := BenchUut7.Slab_Fault_History[0];
   TraceOut_Slab_Fault_History_1[69] := BenchUut7.Slab_Fault_History[1];
   TraceOut_Slab_Fault_History_2[69] := BenchUut7.Slab_Fault_History[2];
   TraceOut_Slab_Fault_History_3[69] := BenchUut7.Slab_Fault_History[3];
   TraceOut_Slab_Fault_History_4[69] := BenchUut7.Slab_Fault_History[4];
   BenchCalls := BenchCalls + 1;
   BenchStep := BenchStep + 1;
  END_IF;
 END_CASE;
 END_IF;
 IF BenchStep >= 70 THEN BenchDone := TRUE; END_IF;
END_IF;
END_PROGRAM
